(* IEC 61131-3 sources: daoli-st-library/DL_Device (part 12) *)

(* ---- FB_DL_AnalogTransmitter.st ---- *)
(*==============================================================================
 * 组件名称 (Component)  : FB_DL_AnalogTransmitter
 * 所属子库 (Sublibrary) : DL_Device
 * 当前版本 (Version)    : 1.0.0
 * 兼容性   (Platform)   : CODESYS 3.5 / TwinCAT 3 / 汇川 InoProShop / Machine Expert
 *                         仅依赖 Standard.library，零厂商方言
 * 分类     (Category)   : 设备信号处理功能块（Function Block，实现 I_DL_AnalogSensor）
 * 功能简述 (Function)   : NAMUR NE43 语义模拟量变送器处理块。在原始物理域
 *                         （mA/0..10V，由调用方约定）执行四段诊断：故障门限外
 *                         断线（方向可配置）、欠量程段、有效测量域、超量程段，
 *                         0 域附近判回路开路；内嵌滑动平均滤波与线性标定；
 *                         故障态保持末次有效工程量；HH/H/L/LL 四级报警在
 *                         有效与欠/超量程段照常计算、故障态全部保持。
 * 接口实现 (Implements) : I_DL_AnalogSensor（属性 fValue/eQuality/bAlarmHH/
 *                         bAlarmH/bAlarmL/bAlarmLL/uErrorId，全部在本文件
 *                         尾部落地）
 * 开源溯源 (Origin)     : 来源标签 namur-ne43（RAW_NOTES_R5 S-5：NAMUR NE43
 *                         信号电平域，公开推荐实践，多来源交叉印证——有效
 *                         测量域 3.8~20.5 mA、故障域 <3.6 / >21 mA、0 mA =
 *                         回路断线、断线诊断须在原始域而非工程量域判定、
 *                         故障方向可配置、超量程标记而非剔除；仅借鉴公开
 *                         标准语义，欠/超量程段以故障门限与量程端点为界
 *                         （默认 4~20 mA 组态下对应 NE43 3.8/20.5 mA 有效
 *                         域界语义），不硬编码，clean-room 未复制任何源码行）。
 * 红线自检 (Redline)    : R1 零全局变量表/外部变量引用 ✓｜R2 零物理 IO 地址 ✓
 *                         R3 纯 IEC 61131-3 ✓｜R4 防除零/防越界/NaN 自比防御 ✓
 *                         R5 全变量中英双语同行注释 ✓｜R6 质量分级判定含
 *                         ELSE 兜底链 ✓｜R7 滤波实例主体无条件刷新（无定时
 *                         器/边缘实例，滤波为纯算术递推）✓
 * 公约遵循 (Convention) : 0.1 首扫判据 IF bTrack OR (NOT _bInit)，跟踪脉冲
 *                         运行中途插入时重置滤波缓冲与保持值。
 *                         0.6 量程对调自修复：对调后继续计算不中断。
 *                         0.8 全部 REAL 输入 fX <> fX 检测，默认值先赋。
 *                         0.7 故障码段位 16#0003_xxxx：【故障级】0003_0210
 *                         NE43 故障态（断线/开路/非有限输入，R15 锁存语义
 *                         由质量位持续标注，原始恢复后自动解除并保持值
 *                         重新跟随）；【信息级】0003_0102 量程对调自修复 /
 *                         0003_0103 欠/超量程提示 / 0003_0104 原始量程跨度
 *                         退化回退（仅写 uErrorId，不设任何故障位，0.2）。
 * 偏离留档 (Deviation)  : 依 R11 头注释留档，共 4 条：
 *                         ① fFilterTC 已按规格 1.6 定稿删除，由 uFilterWindow
 *                           : USINT := 8 滑动平均窗口替代（规格内定稿）。
 *                         ② 引脚表未列 bTrack，为落实 0.1 首扫/跟踪范式与
 *                           "运行中途插入跟踪脉冲"验收向量新增 IN 引脚。
 *                         ③ FC_DL_LinearScale / FB_DL_MovingAverage 本轮
 *                           尚未入库，标定与滤波在本文件内联等价实现（含
 *                           防除零与窗口钳位），两件入库后可无缝外移。
 *                         ④ 对调自修复码 0.6 原文为 16#0001_0001，依 0.7
 *                           段位分配 DL_Device 族取信息级 0003_0102；新增
 *                           0003_0103/0003_0104 按 0.7 之 01xx 信息段顺延。
 * 修订历史 (Revision)   :
 *   2026-11-15  v1.0.0  首版入库（R5 轮 · DL_Device 开库）
 *============================================================================*)

(*-----------------------------------------------------------------------------
 * 枚举: E_DL_BreakDir（归属 FB_DL_AnalogTransmitter，与其同文件）
 * 含义: 断线故障方向配置，由变送器实际 Downscale/Upscale 组态决定；
 *       只判配置方向，另一方向的越限不误报为断线（S-5 提取点②）。
 *----------------------------------------------------------------------------*)
TYPE E_DL_BreakDir :
(
    eLow  := 0,    // 低断方向（Downscale）：原始值低于故障下门限判断线 / Downscale direction, raw below low fault threshold means wire break
    eHigh := 1     // 高断方向（Upscale）：原始值高于故障上门限判断线 / Upscale direction, raw above high fault threshold means wire break
) USINT;
END_TYPE

(*==============================================================================
 * 功能块主体
 *============================================================================*)
FUNCTION_BLOCK FB_DL_AnalogTransmitter IMPLEMENTS I_DL_AnalogSensor
VAR_INPUT
    fRawInput      : REAL;              // 原始输入（Raw input），已线性化的 mA/0..10V 物理域值，单位由调用方约定 / Raw physical-domain input, unit per caller config
    fRawLow        : REAL;              // 原始域量程下限（Raw span low），如 4.0 mA；对调自修复 / Raw span low endpoint, swap self-repair
    fRawHigh       : REAL;              // 原始域量程上限（Raw span high），如 20.0 mA；对调自修复 / Raw span high endpoint, swap self-repair
    fEuLow         : REAL;              // 工程量程下限（Engineering span low），如 0.0 [%] 或 [kPa] / Engineering span low endpoint
    fEuHigh        : REAL;              // 工程量程上限（Engineering span high），如 100.0 [%] 或 [kPa] / Engineering span high endpoint
    eBreakDirection: E_DL_BreakDir := E_DL_BreakDir.eLow; // 断线故障方向（Break direction），eLow=低断 / eHigh=高通，按变送器组态 / Break direction per transmitter config
    fFaultLow      : REAL := 3.6;       // NE43 故障下门限（NE43 low fault threshold），默认 3.6（原始域）/ Low fault threshold in raw domain
    fFaultHigh     : REAL := 21.0;      // NE43 故障上门限（NE43 high fault threshold），默认 21.0（原始域）/ High fault threshold in raw domain
    uFilterWindow  : USINT := 8;        // 滑动平均窗口（Moving-average window），规格定稿替代时间常数引脚，1=直通 / Moving-average window, 1 = pass-through
    bEnableFilter  : BOOL := TRUE;      // 使能滑动平均滤波（Enable moving-average filter），FALSE=直通 / FALSE bypasses filtering
    fAlarmHH       : REAL;              // 上上限报警门限（High-high alarm limit），量纲=工程量 / High-high limit in engineering unit, 非数=禁用 / NaN disables
    fAlarmH        : REAL;              // 上限报警门限（High alarm limit），量纲=工程量，非数=禁用 / High limit in engineering unit, NaN disables
    fAlarmL        : REAL;              // 下限报警门限（Low alarm limit），量纲=工程量，非数=禁用 / Low limit in engineering unit, NaN disables
    fAlarmLL       : REAL;              // 下下限报警门限（Low-low alarm limit），量纲=工程量，非数=禁用 / Low-low limit in engineering unit, NaN disables
    bTrack         : BOOL;              // 跟踪脉冲（Track pulse），上升语义电平：TRUE 拍重置滤波与保持值（R11 偏离新增，见头注释②）/ Track pulse re-primes filter and hold value
END_VAR

VAR_OUTPUT
    fValue         : REAL;              // 工程量当前值（Current engineering value），故障态保持末次有效值 / Holds last good value in fault
    eQuality       : E_DL_SignalQuality; // 信号质量分级（Signal quality grade），NE43 四段诊断 / NE43 diagnostic grade
    bAlarmHH       : BOOL;              // 上上限报警（High-high alarm），有效及欠/超量程段照常计算 / Computed in good and range-violation segments
    bAlarmH        : BOOL;              // 上限报警（High alarm）/ High alarm
    bAlarmL        : BOOL;              // 下限报警（Low alarm）/ Low alarm
    bAlarmLL       : BOOL;              // 下下限报警（Low-low alarm）/ Low-low alarm
    uErrorId       : UDINT;             // 末次故障码（Last error code），0=无故障，段位 16#0003_xxxx / Last error code, 0 = none
    bWireBreak     : BOOL;              // 断线/开路合并位（Wire break merged flag），含开路 / TRUE on wire break or open loop
    bRangeViol     : BOOL;              // 欠/超量程合并位（Range violation merged flag）/ TRUE on under-range or over-range
END_VAR

VAR
    _bInit         : BOOL := FALSE;     // 首扫初始化标志（First-scan init flag），R19 范式判据成员 / R19 paradigm member
    _fHoldEu       : REAL := 0.0;       // 末次有效工程量（Last good engineering value），保持语义载体 / Hold-semantics carrier
    _fValueOut     : REAL := 0.0;       // 输出镜像寄存（Output mirror register），属性与引脚同源 / Mirror shared by pin and property
    _eQualityInt   : E_DL_SignalQuality := E_DL_SignalQuality.eGood; // 质量分级内部寄存（Internal quality register）/ Internal quality register
    _bAlarmHH      : BOOL;              // 上上限报警内部寄存（Internal high-high alarm register）/ Internal alarm register
    _bAlarmH       : BOOL;              // 上限报警内部寄存（Internal high alarm register）/ Internal alarm register
    _bAlarmL       : BOOL;              // 下限报警内部寄存（Internal low alarm register）/ Internal alarm register
    _bAlarmLL      : BOOL;              // 下下限报警内部寄存（Internal low-low alarm register）/ Internal alarm register
    _uErrorIdInt   : UDINT := 0;        // 故障码内部寄存（Internal error code register）/ Internal error code register
    _bFaultState   : BOOL;              // NE43 故障态标志（NE43 fault state flag），断线/开路/非有限输入 / Fault state on break, open loop or non-finite input
    _fRawLoEff     : REAL;              // 对调修复后量程下限（Repaired span low）/ Repaired raw span low endpoint
    _fRawHiEff     : REAL;              // 对调修复后量程上限（Repaired span high）/ Repaired raw span high endpoint
    _bSwap         : BOOL;              // 本拍发生对调修复（Swap repair occurred this cycle）/ Swap repair occurred flag
    _bSpanDegenerate : BOOL;            // 原始量程跨度退化（Degenerate raw span），近零或非有限 / Span near zero or non-finite
    _fFaultLoEff   : REAL := 3.6;       // 防御后故障下门限（Sanitized low fault threshold）/ Sanitized low fault threshold
    _fFaultHiEff   : REAL := 21.0;      // 防御后故障上门限（Sanitized high fault threshold）/ Sanitized high fault threshold
    _fEuLoEff      : REAL := 0.0;       // 防御后工程下限（Sanitized engineering low）/ Sanitized engineering low
    _fEuHiEff      : REAL := 100.0;     // 防御后工程上限（Sanitized engineering high）/ Sanitized engineering high
    _bValid        : BOOL;              // 原始输入有效（Raw input valid），非有限值为 FALSE / FALSE when input is non-finite
    _fScaleRaw     : REAL;              // 参与标定的原始值（Raw value entering scaling），滤波输出或直通 / Filtered or pass-through raw value
    _fScaledEu     : REAL;              // 本拍标定结果（Scaled result this cycle）/ Scaled engineering result this cycle
    _fRawSpan      : REAL;              // 原始量程跨度（Raw span width）/ Raw span width
    _bFilterActive : BOOL;              // 滤波激活（Filter active），使能且窗口 >= 2 / Active when enabled and window >= 2
    _uWindowEff    : USINT;             // 钳位后有效窗口（Effective clamped window），上限 128 / Effective window clamped to 128
    _uWindowPrev   : USINT;             // 上一拍有效窗口（Previous effective window），变更检测用于缓冲重置 / Previous window for change detection
    _uBufIdx       : UINT;              // 环形缓冲写指针（Ring buffer write index），0..127 / Ring write index 0..127
    _uBufFill      : USINT;             // 有效样本数（Valid sample count），上限=有效窗口 / Valid samples, capped at effective window
    _fBufSum       : REAL := 0.0;       // 窗口样本和（Window sample sum），每拍重算 / Recomputed each cycle
    _fFillR        : REAL := 1.0;       // 样本数实型镜像（Sample count REAL mirror），供安全除法 / REAL mirror of sample count for safe division
    _afBuf         : ARRAY[0..127] OF REAL; // 滑动平均环形缓冲（Moving-average ring buffer），128 槽 / 128-slot ring buffer
    i              : UINT;              // 缓冲遍历循环索引（Buffer traversal loop index）/ Loop index for buffer traversal
    _uRingIdx      : UINT;              // 环形取数临时索引（Ring fetch temp index）/ Temporary ring fetch index
END_VAR

// ============================================================================
// 段 1｜首扫/跟踪初始化（R19 唯一合法范式：IF bTrack OR (NOT _bInit)）
//      First-scan / track initialization (R19 sole legal paradigm)
// ============================================================================
IF bTrack OR (NOT _bInit) THEN
    _uBufIdx   := 0;                          // 写指针归零（Write index reset）
    _uBufFill  := 0;                          // 有效样本清零：滤液从直通逐步重新填充（Samples cleared, filter refills from pass-through）
    _fBufSum   := 0.0;                        // 窗口和清零（Window sum cleared）
    _fHoldEu   := 0.0;                        // 保持值清零，本拍有效样本将立即回填（Hold cleared, refilled by first valid sample）
    _bFaultState := FALSE;                    // 故障态复位（Fault state released）
    _uErrorIdInt := 0;                        // 故障码清零（Error code cleared）
    _eQualityInt := E_DL_SignalQuality.eGood; // 质量复位为良好（Quality reset to good）
    _bInit      := TRUE;                      // 初始化完成（Initialization done）
END_IF

// ============================================================================
// 段 2｜窗口参数钳位与变更检测（防越界：窗口上限 128 槽缓冲）
//      Window clamping and change detection (bounds defense: 128-slot buffer)
// ============================================================================
_uWindowEff := uFilterWindow;                 // 取组态窗口（Take configured window）
IF _uWindowEff > 128 THEN
    _uWindowEff := 128;                       // 超限钳位到缓冲容量（Clamp to buffer capacity）
END_IF
IF _uWindowEff = 0 THEN
    _uWindowEff := 1;                         // 零窗口按单样本直通（Zero window treated as single-sample pass-through）
END_IF
IF _uWindowEff <> _uWindowPrev THEN           // 窗口在线变更（Window changed online）
    _uBufFill := 0;                           // 缓冲判无效重新填充（Invalidate buffer, refill from scratch）
    _uWindowPrev := _uWindowEff;              // 记录新窗口（Record new window）
END_IF
_bFilterActive := bEnableFilter AND (_uWindowEff >= 2); // 窗口 1 视为直通（Window 1 treated as pass-through）

// ============================================================================
// 段 3｜参数防御（0.8：全部 REAL 参数先做非数自比，默认值先赋）+ 0.6 对调自修复
//      Parameter sanitation (0.8 NaN self-compare, defaults first) + 0.6 swap repair
// ============================================================================
_fRawLoEff := fRawLow;                        // 量程下限镜像（Span low mirror）
_fRawHiEff := fRawHigh;                       // 量程上限镜像（Span high mirror）
_fEuLoEff  := fEuLow;                         // 工程下限镜像（Engineering low mirror）
_fEuHiEff  := fEuHigh;                        // 工程上限镜像（Engineering high mirror）
_fFaultLoEff := fFaultLow;                    // 故障下门限镜像（Low fault threshold mirror）
_fFaultHiEff := fFaultHigh;                   // 故障上门限镜像（High fault threshold mirror）

IF _fFaultLoEff <> _fFaultLoEff THEN          // 非数自比检测（NaN self-compare test）
    _fFaultLoEff := 3.6;                      // 回落 NE43 默认下门限（Fallback to NE43 default low）
END_IF
IF _fFaultHiEff <> _fFaultHiEff THEN          // 非数自比检测（NaN self-compare test）
    _fFaultHiEff := 21.0;                     // 回落 NE43 默认上门限（Fallback to NE43 default high）
END_IF
IF _fEuLoEff <> _fEuLoEff THEN                // 非数自比检测（NaN self-compare test）
    _fEuLoEff := 0.0;                         // 回落工程下限默认（Fallback engineering low default）
END_IF
IF _fEuHiEff <> _fEuHiEff THEN                // 非数自比检测（NaN self-compare test）
    _fEuHiEff := 100.0;                       // 回落工程上限默认（Fallback engineering high default）
END_IF

_bSwap := FALSE;                              // 对调标志复位（Swap flag reset）
IF _fRawLoEff > _fRawHiEff THEN               // 参数对自修复判据（Pair swap test, NaN-safe ordering）
    _fRawLoEff := fRawHigh;                   // 下限取原上限（Low takes former high）
    _fRawHiEff := fRawLow;                    // 上限取原下限（High takes former low）
    _bSwap := TRUE;                           // 登记对调修复（Register swap repair, computation continues）
END_IF

// ============================================================================
// 段 4｜非有限输入判定（0.8）与出口默认值先赋（保持语义）
//      Non-finite input test (0.8) and output defaults assigned first (hold)
// ============================================================================
_bValid := (fRawInput = fRawInput);           // 非数自比检测：等号成立即有效（NaN 时自比不等）/ NaN iff self-compare fails, TRUE means valid
_fValueOut := _fHoldEu;                       // 出口默认：保持末次有效值（Default: hold last good value）
_bFaultState := FALSE;                        // 故障态先复位，分级链中重新判定（Fault state preset FALSE, re-decided below）
_eQualityInt := E_DL_SignalQuality.eGood;     // 出口默认质量（Default quality）

// ============================================================================
// 段 5｜NE43 四段质量分级（全部在原始物理域判定，S-5 提取点③；
//       断线只判配置方向，配置外方向不误报）
//      NE43 four-band classification in raw domain, break judged only on
//      the configured direction to avoid false breaks
// ============================================================================

IF NOT _bValid THEN
    _eQualityInt := E_DL_SignalQuality.eOpenLoop;   // 非有限输入按回路开路处理（Non-finite input as open loop）
    _bFaultState := TRUE;                           // 进入故障态（Enter fault state）
ELSIF fRawInput < (_fFaultLoEff * 0.5) THEN
    _eQualityInt := E_DL_SignalQuality.eOpenLoop;   // 0 域附近判开路（0 mA 回路断开）/ Near-zero domain as open loop
    _bFaultState := TRUE;
ELSIF fRawInput < _fFaultLoEff THEN
    IF eBreakDirection = E_DL_BreakDir.eLow THEN
        _eQualityInt := E_DL_SignalQuality.eWireBreakLow; // 配置低断：判断线（Configured downscale: wire break）
        _bFaultState := TRUE;
    ELSE
        _eQualityInt := E_DL_SignalQuality.eUnderRange;   // 配置高通：欠量程段不误报断线（High config: under-range, no false break）
    END_IF
ELSIF fRawInput > _fFaultHiEff THEN
    IF eBreakDirection = E_DL_BreakDir.eHigh THEN
        _eQualityInt := E_DL_SignalQuality.eWireBreakHigh; // 配置高通：判断线（Configured upscale: wire break）
        _bFaultState := TRUE;
    ELSE
        _eQualityInt := E_DL_SignalQuality.eOverRange;     // 配置低断：超量程段不误报断线（Low config: over-range, no false break）
    END_IF
ELSIF fRawInput < _fRawLoEff THEN
    _eQualityInt := E_DL_SignalQuality.eUnderRange;   // 欠量程段（如 3.6~4.0 mA）标记不剔除（Under-range marked, not discarded）
ELSIF fRawInput > _fRawHiEff THEN
    _eQualityInt := E_DL_SignalQuality.eOverRange;    // 超量程段（如 20.0~21.0 mA）标记不剔除（Over-range marked, not discarded）
ELSE
    _eQualityInt := E_DL_SignalQuality.eGood;         // 有效测量域（Valid measurement span）
END_IF

// ============================================================================
// 段 6｜滑动平均滤波（仅有效拍推入缓冲，故障拍不污染窗口）+ 线性标定
//      Moving-average filter (push only on valid cycles) + linear scaling
// ============================================================================
IF _bFaultState THEN
    _fScaleRaw := fRawInput;                  // 故障拍标定值不使用（Unused in fault cycles, hold applies）
ELSE
    IF _bFilterActive THEN
        _afBuf[_uBufIdx] := fRawInput;        // 写入环形槽（Write ring slot, index < 128 by MOD）
        _uBufIdx := (_uBufIdx + 1) MOD 128;   // 写指针循环推进（Advance write index cyclically）
        IF _uBufFill < _uWindowEff THEN
            _uBufFill := _uBufFill + 1;       // 未满则递增有效样本（Increment fill until window reached）
        END_IF
        _fBufSum := 0.0;                      // 每拍重算窗口和（Recompute window sum each cycle）
        FOR i := 1 TO _uBufFill DO            // 固定界循环，无死循环风险（Bounded loop, no deadlock risk）
            _uRingIdx := (_uBufIdx + 128 - i) MOD 128; // 倒序取最近样本槽（Fetch latest slots in reverse order）
            _fBufSum := _fBufSum + _afBuf[_uRingIdx];  // 累加窗口样本（Accumulate window sample）
        END_FOR
        _fFillR := _uBufFill;                 // 样本数实型镜像（Sample count as REAL）
        IF _fFillR > 0.5 THEN
            _fScaleRaw := _fBufSum / _fFillR; // 窗口均值（Window mean, divisor proven >= 1）
        ELSE
            _fScaleRaw := fRawInput;          // 防除零回退直通（Divide-by-zero fallback to pass-through）
        END_IF
    ELSE
        _fScaleRaw := fRawInput;              // 滤波禁用直通（Filter disabled, pass-through）
    END_IF

    // 线性标定（内联实现，偏离留档③；除零与退化双重防御）
    _fRawSpan := _fRawHiEff - _fRawLoEff;     // 原始量程跨度（Raw span width）
    _bSpanDegenerate := (_fRawSpan <> _fRawSpan) OR (ABS(_fRawSpan) < 1E-9); // 非数或近零判退化（Degenerate on NaN or near-zero）
    IF _bSpanDegenerate THEN
        _fScaledEu := _fEuLoEff;              // 退化回退工程下限（Degenerate fallback to engineering low）
    ELSE
        _fScaledEu := _fEuLoEff + (_fScaleRaw - _fRawLoEff) * (_fEuHiEff - _fEuLoEff) / _fRawSpan; // 线性插值（Linear interpolation, denominator proven non-zero）
    END_IF
    _fValueOut := _fScaledEu;                 // 有效拍输出跟随（Output follows on valid cycles）
    _fHoldEu   := _fScaledEu;                 // 更新保持载体（Update hold carrier）
END_IF

// ============================================================================
// 段 7｜四级报警计算（有效与欠/超量程段照常计算；故障态全部保持；
//       门限为非数时该级视为未组态不报警——0.8 防御）
//      Four-level alarms (computed in good and range segments, held in
//      fault; NaN threshold disables that level)
// ============================================================================
IF NOT _bFaultState THEN
    IF fAlarmHH = fAlarmHH THEN
        _bAlarmHH := (_fValueOut >= fAlarmHH); // 上上限判定（High-high evaluation）
    ELSE
        _bAlarmHH := FALSE;                    // 门限非数=该级禁用（NaN limit disables level）
    END_IF
    IF fAlarmH = fAlarmH THEN
        _bAlarmH := (_fValueOut >= fAlarmH);   // 上限判定（High evaluation）
    ELSE
        _bAlarmH := FALSE;                     // 门限非数=该级禁用（NaN limit disables level）
    END_IF
    IF fAlarmL = fAlarmL THEN
        _bAlarmL := (_fValueOut <= fAlarmL);   // 下限判定（Low evaluation）
    ELSE
        _bAlarmL := FALSE;                     // 门限非数=该级禁用（NaN limit disables level）
    END_IF
    IF fAlarmLL = fAlarmLL THEN
        _bAlarmLL := (_fValueOut <= fAlarmLL); // 下下限判定（Low-low evaluation）
    ELSE
        _bAlarmLL := FALSE;                    // 门限非数=该级禁用（NaN limit disables level）
    END_IF
END_IF // 故障态不进入本段，四级报警输出自动保持上一拍值（Fault cycles skip this block, alarms held）

// ============================================================================
// 段 8｜故障码优先级链与合并位派生（信息级仅写 uErrorId，0.2 公约）
//      Error-code priority chain and merged flag derivation (info codes only)
// ============================================================================
IF _bFaultState THEN
    _uErrorIdInt := 16#0003_0210;             // 0003_0210 NE43 故障态（断线/开路/非有限输入）【故障级】/ NE43 fault state, fault level
ELSIF (_eQualityInt = E_DL_SignalQuality.eUnderRange) OR (_eQualityInt = E_DL_SignalQuality.eOverRange) THEN
    _uErrorIdInt := 16#0003_0103;             // 0003_0103 欠/超量程提示【信息级】/ Range violation hint, info level
ELSIF _bSwap THEN
    _uErrorIdInt := 16#0003_0102;             // 0003_0102 量程对调自修复【信息级】（0.6 公约，段位依 0.7 归 DL_Device 信息段）/ Swap self-repair, info level
ELSIF _bSpanDegenerate THEN
    _uErrorIdInt := 16#0003_0104;             // 0003_0104 原始量程跨度退化回退【信息级】/ Degenerate span fallback, info level
ELSE
    _uErrorIdInt := 0;                        // 无故障无提示（No fault, no hint）
END_IF

// ============================================================================
// 段 9｜引脚映射（属性与引脚同源于内部镜像，避免同名遮蔽）
//      Pin mapping (pin and property share internal mirrors, no shadowing)
// ============================================================================
fValue     := _fValueOut;                     // 工程量输出（Engineering value output）
eQuality   := _eQualityInt;                   // 质量分级输出（Quality output）
bAlarmHH   := _bAlarmHH;                      // 上上限输出（High-high output）
bAlarmH    := _bAlarmH;                       // 上限输出（High output）
bAlarmL    := _bAlarmL;                       // 下限输出（Low output）
bAlarmLL   := _bAlarmLL;                      // 下下限输出（Low-low output）
uErrorId   := _uErrorIdInt;                   // 故障码输出（Error code output）
bWireBreak := (_eQualityInt = E_DL_SignalQuality.eWireBreakLow)
          OR (_eQualityInt = E_DL_SignalQuality.eWireBreakHigh)
          OR (_eQualityInt = E_DL_SignalQuality.eOpenLoop);            // 断线/开路合并位（Break/open merged flag）
bRangeViol := (_eQualityInt = E_DL_SignalQuality.eUnderRange)
          OR (_eQualityInt = E_DL_SignalQuality.eOverRange);           // 欠/超量程合并位（Range violation merged flag）

(*------------------------------------------------------------------------------
 * 属性: fValue（GET）—— 工程量当前值（故障态保持末次有效值）。
 *      Property fValue (GET) - current engineering value, holds last good in fault.
 *------------------------------------------------------------------------------*)
PROPERTY fValue : REAL
fValue := _fValueOut;         // 返回输出镜像（Return output mirror）

(*------------------------------------------------------------------------------
 * 属性: eQuality（GET）—— 信号质量分级（NE43 四段诊断结果）。
 *      Property eQuality (GET) - signal quality grade per NE43 diagnostics.
 *------------------------------------------------------------------------------*)
PROPERTY eQuality : E_DL_SignalQuality
eQuality := _eQualityInt;     // 返回质量镜像（Return quality mirror）

(*------------------------------------------------------------------------------
 * 属性: bAlarmHH（GET）—— 上上限报警位。
 *      Property bAlarmHH (GET) - high-high alarm bit.
 *------------------------------------------------------------------------------*)
PROPERTY bAlarmHH : BOOL
bAlarmHH := _bAlarmHH;        // 返回上上限镜像（Return high-high mirror）

(*------------------------------------------------------------------------------
 * 属性: bAlarmH（GET）—— 上限报警位。
 *      Property bAlarmH (GET) - high alarm bit.
 *------------------------------------------------------------------------------*)
PROPERTY bAlarmH : BOOL
bAlarmH := _bAlarmH;          // 返回上限镜像（Return high mirror）

(*------------------------------------------------------------------------------
 * 属性: bAlarmL（GET）—— 下限报警位。
 *      Property bAlarmL (GET) - low alarm bit.
 *------------------------------------------------------------------------------*)
PROPERTY bAlarmL : BOOL
bAlarmL := _bAlarmL;          // 返回下限镜像（Return low mirror）

(*------------------------------------------------------------------------------
 * 属性: bAlarmLL（GET）—— 下下限报警位。
 *      Property bAlarmLL (GET) - low-low alarm bit.
 *------------------------------------------------------------------------------*)
PROPERTY bAlarmLL : BOOL
bAlarmLL := _bAlarmLL;        // 返回下下限镜像（Return low-low mirror）

(*------------------------------------------------------------------------------
 * 属性: uErrorId（GET）—— 末次故障码（0=无故障）。
 *      Property uErrorId (GET) - last error code (0 = none).
 *------------------------------------------------------------------------------*)
PROPERTY uErrorId : UDINT
uErrorId := _uErrorIdInt;     // 返回故障码镜像（Return error code mirror）
END_FUNCTION_BLOCK

(* ---- FB_DL_AnalogValve.st ---- *)
(*==============================================================================
 * 组件名称 (Component)  : FB_DL_AnalogValve
 * 所属子库 (Sublibrary) : DL_Device
 * 当前版本 (Version)    : 1.0.1
 * 兼容性   (Platform)   : CODESYS 3.5 / TwinCAT 3 / 汇川 InoProShop / Machine Expert
 *                         仅依赖 Standard.library（TON / R_TRIG），零厂商方言
 * 分类     (Category)   : 设备执行器功能块（Function Block，实现 I_DL_ProportionalValve）
 * 功能简述 (Function)   : 模拟量比例阀指令整形与诊断功能块（不含阀位闭环，
 *                         闭环由驱动器/上层 PID 完成，本块职责单一）。
 *                         透传+补偿链：设定钳位 [0,100] → 零点死区补偿
 *                         （防阀芯微抖）→ 限幅域映射 → 阀位指令输出；
 *                         偏差报警延时确认（瞬时型每拍重算，恢复自动清）；
 *                         非有限值反馈锁存保持末次有效值；限幅域对调
 *                         自修复；状态机 E_DL_ValveState + CASE + ELSE
 *                         兜底。
 * 接口实现 (Implements) : I_DL_ProportionalValve。接口 OUT 列同名成员
 *                         （eState/fPosCmd/fPosFeedback/bDeviationAlarm/
 *                         bFault/uErrorId）按 R22 以只读 PROPERTY GET
 *                         承载（内部镜像同源；fPosFeedback 为 IN 引脚与
 *                         接口属性双形式暴露，沿用库级既有先例），非接口
 *                         成员 fPosOutput 保留 VAR_OUTPUT；方法
 *                         SetPosition/CmdStop/CmdReset 全部在本文件尾部
 *                         落地。
 * 开源溯源 (Origin)     : 来源标签 lbp-basic-process / lbp-device
 *                         （RAW_NOTES_R6 S-1：比例阀指令整形链（钳位-死区
 *                         补偿-限幅域映射）、偏差延时报警、限幅域端点组态
 *                         等行业公知工程惯例，公开教学资料，仅借鉴通用
 *                         工程语义；状态机、整形链实现、故障码按本库红线
 *                         独立设计，clean-room 未复制源码）。
 * 红线自检 (Redline)    : R1 零全局变量表/外部变量引用 ✓｜R2 零物理 IO 地址 ✓
 *                         R3 纯 IEC 61131-3 ✓｜R4 防除零/防越界/非有限值
 *                         防御/浮点容差比较 ✓｜R5 全变量中英双语同行注释 ✓
 *                         R6 ENUM+CASE+ELSE ✓｜R7 两个定时器/边缘实例主体
 *                         最前部无条件刷新 ✓
 * 公约遵循 (Convention) : 0.1/R23 本块为逐拍组合整形链（设定→钳位→死区→
 *                         映射，全部由实时输入重算自校正），无积分/滤波类
 *                         需要首扫初始化的连续量驻留状态，免首扫（无
 *                         bInit 标志）；时间基准按公约 0.5 采用 TON 延时
 *                         引脚（偏差确认），无采样周期类连续量语义。
 *                         0.6 限幅域对调自修复：fOutMin > fOutMax 时对调
 *                         + 置信息级码 + 继续计算不中断。
 *                         0.7 故障码段位 16#0003_xxxx：【故障级】0003_0260
 *                         阀位反馈信号无效 / 0003_0261 非法状态，R15 锁存
 *                         仅复位可清；【信息级】0003_0108 设定值钳位 /
 *                         0003_0109 输出限幅域对调自修复 / 0003_0112 偏差
 *                         报警激活（瞬时型每拍重算，0.15；不进 bFault）。
 * 偏离留档 (Deviation)  : 依 R11 头注释留档，共 1 条：
 *                         ① 信息级码：规格原分配 0003_0105/0106，经与子库
 *                           VERSION.md 故障码表核对，R5 已占用 0102~0104
 *                           （AnalogTransmitter），且 0106/0107 已由本轮
 *                           变频器块顺延占用（0105 经终审裁定空置：重启抑
 *                           制拒绝统一沿用 DolMotor 既有语义码位 0208），
 *                           依公约 0.7 冲突顺延：设定值钳位 → 0108、限幅
 *                           域对调 → 0109；偏差报警激活为新码位，顺延分配
 *                           0112。
 * 修订历史 (Revision)   :
 *   2026-11-15  v1.0.0  首版入库（R6 轮 · DL_Device 阀门/驱动族深化）
 *   2026-11-15  v1.0.1  终审修复【工程语义级】限幅域对调穿透：原实现对调时
 *                       直读原始引脚（fOutMin/fOutMax），混合非数组态下
 *                       （如下端非数+上端负值）会把未防御的 NaN 带回生效
 *                       域并经映射链输出 NaN 阀位指令且不带故障码。修法：
 *                       对调改为经中间变量交换已防御的生效值。引脚契约
 *                       零变更。
 *============================================================================*)
FUNCTION_BLOCK FB_DL_AnalogValve IMPLEMENTS I_DL_ProportionalValve
VAR_INPUT
    fPosSetpoint     : REAL;            // 阀位设定（Position setpoint）[%]，0..100，越界钳位信息级 / Position setpoint [%], clamped with info code
    fPosFeedback     : REAL;            // 阀位反馈（Position feedback）[%]，0..100，来自阀位变送器；非有限值防御 / Position feedback [%] from transmitter, non-finite defended
    fZeroDeadband    : REAL := 0.5;     // 零点死区补偿（Zero deadband compensation）[%]，输出小于此值钳为 0 防阀芯微抖 / Zero deadband [%], output below clamped to zero
    fDeviationLimit  : REAL := 5.0;     // 偏差报警门限（Deviation limit）[%]，默认 5.0 / Deviation alarm limit [%], default 5.0
    tDeviationDelay  : TIME := T#10S;   // 偏差报警确认延时（Deviation delay），防动态调节过程误报 / Deviation confirmation delay against dynamic transients
    fOutMin          : REAL := 0.0;     // 输出限幅域下端点（Output span low endpoint）[%]，对调自修复 / Output span low endpoint, swap self-repair
    fOutMax          : REAL := 100.0;   // 输出限幅域上端点（Output span high endpoint）[%]，对调自修复 / Output span high endpoint, swap self-repair
    bEnable          : BOOL;            // 调节使能（Modulating enable），FALSE 时输出冻结保持 / Modulating enable, FALSE freezes output hold
    bReset           : BOOL;            // 故障复位（Fault reset），上升沿生效 / Fault reset, rising edge effective
END_VAR

VAR_OUTPUT
    fPosOutput : REAL;                  // 阀位指令输出（Position output）[%]，死区补偿+限幅域映射后，量纲=限幅域（R20）/ Shaped position output [%], span of limit domain
END_VAR

VAR
    _eState        : E_DL_ValveState := E_DL_ValveState.eIdle; // 内部状态机步序（Internal state step），外部经属性只读 / Internal state, read-only via property
    _bFaultLatch   : BOOL;              // 故障锁存标志（Fault latch flag），仅复位清除 / Fault latch flag, cleared only by reset
    _uErrorIdInt   : UDINT;             // 故障级码内部寄存（Internal fault-code register） / Internal fault-level code register
    _uInfoCode     : UDINT;             // 本拍信息级码（Info code this cycle），瞬时型每拍重算（0.15）/ Transient info code recomputed each cycle
    _bHoldLatch    : BOOL;              // 输出冻结锁存（Output freeze latch），CmdStop 置位 / Output freeze latch set by CmdStop
    _bPendReset    : BOOL;              // 方法复位请求（Method reset request），由 CmdReset 置位 / Method reset request set by CmdReset
    _bClampOccur   : BOOL;              // 本拍设定值钳位发生（Setpoint clamp occurred this cycle）/ Setpoint clamp occurred flag
    _fPosMethVal   : REAL;              // 方法阀位设定值（Method position value）[%] / Position value set via method
    _bPosMethAct   : BOOL;              // 方法阀位设定激活（Method position active），激活后覆盖引脚 / Method position active, overrides pin
    _fPosFbHold    : REAL := 0.0;       // 末次有效阀位反馈（Last valid position feedback）[%]，保持载体 / Last valid feedback hold carrier
    _fPosCmdEff    : REAL := 0.0;       // 钳位+死区后生效阀位指令（Effective command after clamp and deadband）[%] / Effective command [%]
    _fPosOutHold   : REAL := 0.0;       // 输出保持载体（Output hold carrier）[%]，冻结/故障态保持 / Output hold carrier [%]
    _fOutMinEff    : REAL := 0.0;       // 对调修复后限幅域下端（Repaired span low endpoint）[%] / Repaired span low endpoint
    _fOutMaxEff    : REAL := 100.0;     // 对调修复后限幅域上端（Repaired span high endpoint）[%] / Repaired span high endpoint
    _fZeroDbEff    : REAL := 0.5;       // 防御后死区（Sanitized deadband）[%]，非数/负值钳零 / Sanitized deadband, NaN or negative clamped to zero
    _fDevLimEff    : REAL := 5.0;       // 防御后偏差门限（Sanitized deviation limit）[%] / Sanitized deviation limit
    _bSpanSwap     : BOOL;              // 本拍限幅域对调修复（Span swap repair this cycle）/ Span swap repair occurred flag
    _fSpanTmp      : REAL;              // 对调交换中间变量（Swap temp carrier）[%]，生效域已防御值 / Swap temp for sanitized span values
    _bSpanDegenerate : BOOL;            // 限幅域跨度退化（Degenerate span），近零或非有限 / Span degenerate on near-zero or NaN
    _bFbValid      : BOOL;              // 本拍反馈有效性（Feedback validity this cycle），非有限值为 FALSE / FALSE when feedback non-finite
    _bDevRaw       : BOOL;              // 偏差越限原始判据（Raw deviation-exceed test）/ Raw deviation exceed flag
    _bDeviationAct : BOOL;              // 偏差报警激活中（Deviation alarm active），延时确认后 / Deviation alarm active after confirmation delay
    _fbTrigReset   : R_TRIG;            // 引脚复位上升沿（Pin reset edge）/ Pin reset rising edge
    _fbTonDev      : TON;               // 偏差报警确认延时定时器（Deviation confirmation timer）/ Deviation confirmation timer
END_VAR

METHOD SetPosition : BOOL
VAR_INPUT
    fPos : REAL; // 阀位设定值（Position value）[%]，域 0..100 / Position value [%], range 0..100
END_VAR
IF _bFaultLatch OR (_eState = E_DL_ValveState.eFault) THEN
    SetPosition := FALSE;     // 故障态拒绝（Rejected in fault state）
ELSIF (fPos <> fPos) OR (fPos < 0.0) OR (fPos > 100.0) THEN
    SetPosition := FALSE;     // 非数或越域拒绝（Rejected on NaN or out of range）
ELSE
    _fPosMethVal := fPos;     // 登记方法设定值（Register method position value）
    _bPosMethAct := TRUE;     // 激活方法设定通道（Activate method source channel）
    _bHoldLatch  := FALSE;    // 设定即解除输出冻结（Set releases output freeze）
    SetPosition := TRUE;      // 受理成功（Accepted）
END_IF

(*------------------------------------------------------------------------------
 * 方法: CmdStop —— 冻结输出保持当前阀位，直至下次设定或使能撤除。
 *      Method CmdStop - freeze output until next set or enable drop.
 *------------------------------------------------------------------------------*)
    END_METHOD

METHOD CmdStop : BOOL
VAR_INPUT
END_VAR
IF _bFaultLatch OR (_eState = E_DL_ValveState.eFault) THEN
    CmdStop := FALSE;         // 故障态拒绝（Rejected in fault state）
ELSE
    _bHoldLatch := TRUE;      // 登记冻结锁存，主体状态机消化（Register freeze latch, consumed by body）
    CmdStop := TRUE;          // 受理成功（Accepted）
END_IF

(*------------------------------------------------------------------------------
 * 方法: CmdReset —— 复位故障，返回是否可复位（存在锁存故障时为 TRUE）。
 *      Method CmdReset - reset fault, returns TRUE only when a latch exists.
 *------------------------------------------------------------------------------*)
    END_METHOD

METHOD CmdReset : BOOL
VAR_INPUT
END_VAR
IF _bFaultLatch OR (_eState = E_DL_ValveState.eFault) THEN
    _bPendReset := TRUE;      // 登记复位请求，主体状态机消化（Register reset request, consumed by body）
    CmdReset := TRUE;         // 可复位（Resettable）
ELSE
    CmdReset := FALSE;        // 无故障可复位（Nothing to reset）
END_IF

(*------------------------------------------------------------------------------
 * 属性: eState（GET）—— 当前状态机状态只读视图。
 *      Property eState (GET) - read-only view of the current state machine state.
 *------------------------------------------------------------------------------*)
    END_METHOD

// ============================================================================
// 段 1｜定时器与边缘检测实例无条件周期刷新（R7：严禁置于 IF/CASE 分支内）
//      Unconditional per-cycle refresh of all timer and edge instances (R7)
// ============================================================================
_fbTrigReset(CLK := bReset);
_bDevRaw := (_eState = E_DL_ValveState.eModulating) AND (ABS(_fPosCmdEff - _fPosFbHold) > _fDevLimEff); // 偏差原始判据（Raw deviation test）
_fbTonDev(IN := _bDevRaw, PT := tDeviationDelay); // 延时确认防动态调节误报（Delay confirmation against dynamics）

// ============================================================================
// 段 2｜参数防御（0.8：非数自比检测，默认值先赋）+ 0.6 限幅域对调自修复
//      Parameter sanitation (0.8 NaN self-compare) + 0.6 span swap repair
// ============================================================================
_uInfoCode := 0;                      // 本拍信息级码先归零，事件段重算（Info code preset zero, recomputed in event chain）
_bClampOccur := FALSE;                // 钳位标志复位（Clamp flag reset）
_fZeroDbEff := fZeroDeadband;         // 死区镜像（Deadband mirror）
IF _fZeroDbEff <> _fZeroDbEff THEN    // 非数自比检测（NaN self-compare test）
    _fZeroDbEff := 0.0;               // 非数死区钳零禁用补偿（NaN deadband clamped to zero, compensation disabled）
END_IF
IF _fZeroDbEff < 0.0 THEN
    _fZeroDbEff := 0.0;               // 负死区钳零（Negative deadband clamped to zero）
END_IF
_fDevLimEff := fDeviationLimit;       // 偏差门限镜像（Deviation limit mirror）
IF _fDevLimEff <> _fDevLimEff THEN    // 非数自比检测（NaN self-compare test）
    _fDevLimEff := 5.0;               // 回落默认门限（Fallback to default limit）
END_IF
IF _fDevLimEff < 0.0 THEN
    _fDevLimEff := ABS(_fDevLimEff);  // 负门限取绝对值保持报警有效（Negative limit made absolute, alarm stays valid）
END_IF

_fOutMinEff := fOutMin;               // 限幅域下端镜像（Span low mirror）
_fOutMaxEff := fOutMax;               // 限幅域上端镜像（Span high mirror）
IF _fOutMinEff <> _fOutMinEff THEN    // 非数自比检测（NaN self-compare test）
    _fOutMinEff := 0.0;               // 回落下端默认（Fallback to default low）
END_IF
IF _fOutMaxEff <> _fOutMaxEff THEN    // 非数自比检测（NaN self-compare test）
    _fOutMaxEff := 100.0;             // 回落上端默认（Fallback to default high）
END_IF
_bSpanSwap := FALSE;                  // 对调标志复位（Swap flag reset）
IF _fOutMinEff > _fOutMaxEff THEN     // 参数对自修复判据（Pair swap test）
    _fSpanTmp     := _fOutMinEff;     // 对调经已防御的生效值交换（中间变量，防原始引脚
    _fOutMinEff   := _fOutMaxEff;     // 非有限值穿透——若直读原始引脚，混合非数组态
    _fOutMaxEff   := _fSpanTmp;       // 会把 NaN 带回生效域，终审修复）
    _bSpanSwap := TRUE;               // 登记对调修复，继续计算不中断（Register swap repair, computation continues）
END_IF

// ============================================================================
// 段 3｜阀位反馈有效性全局监视（优先级最高，故障级锁存保持末次有效值）
//      Position feedback validity global monitor (highest priority, latched)
// ============================================================================
_bFbValid := (fPosFeedback = fPosFeedback); // 非数自比检测：等号成立即有效（NaN iff self-compare fails）
IF _bFbValid THEN
    _fPosFbHold := fPosFeedback;      // 更新末次有效反馈（Update last valid feedback）
ELSE
    _bFaultLatch := TRUE;             // 反馈失效锁存（Feedback loss latch）
    _uErrorIdInt := 16#0003_0260;     // 0003_0260 阀位反馈信号无效【故障级】/ Position feedback invalid, fault level
    _eState      := E_DL_ValveState.eFault; // 强制故障态（Force fault state）
END_IF

// ============================================================================
// 段 4｜指令整形链：来源选择 → 钳位 [0,100] → 零点死区补偿
//      Command shaping chain: source select → clamp [0,100] → zero deadband
// ============================================================================
IF _bPosMethAct THEN
    _fPosCmdEff := _fPosMethVal;      // 方法设定覆盖引脚（Method value overrides pin）
ELSE
    _fPosCmdEff := fPosSetpoint;      // 引脚设定（Pin setpoint）
END_IF
IF _fPosCmdEff <> _fPosCmdEff THEN    // 非数自比检测（NaN self-compare test）
    _fPosCmdEff := 0.0;               // 非数设定回零（NaN setpoint falls back to zero）
END_IF
IF _fPosCmdEff < 0.0 THEN
    _fPosCmdEff := 0.0;               // 下限钳位（Clamped to low bound）
    _bClampOccur := TRUE;             // 登记钳位事件（Register clamp event）
END_IF
IF _fPosCmdEff > 100.0 THEN
    _fPosCmdEff := 100.0;             // 上限钳位（Clamped to high bound）
    _bClampOccur := TRUE;             // 登记钳位事件（Register clamp event）
END_IF
IF ABS(_fPosCmdEff) < _fZeroDbEff THEN
    _fPosCmdEff := 0.0;               // 零点死区补偿：近零指令钳为 0 防阀芯微抖（Zero deadband: near-zero command clamped to zero）
END_IF

// ============================================================================
// 段 5｜核心状态机（ENUM + CASE，含 ELSE 非法状态兜底）
//      Core state machine (ENUM + CASE with ELSE illegal-state fallback)
// ============================================================================
IF _bFaultLatch OR (_eState = E_DL_ValveState.eFault) THEN
    CASE _eState OF
        E_DL_ValveState.eFault: // 故障锁存态：输出冻结保持，仅复位可退出
            IF _fbTrigReset.Q OR _bPendReset THEN
                _bPendReset  := FALSE;            // 消费复位请求（Consume reset request）
                _bFaultLatch := FALSE;            // 解除锁存（Release latch）
                _uErrorIdInt := 0;                // 故障码清零（Error code cleared）
                _bHoldLatch  := FALSE;            // 复位同时解除冻结（Freeze released on reset）
                _eState      := E_DL_ValveState.eIdle; // 回空闲态（Back to idle）
            END_IF
        ELSE // 锁存标志与状态不一致兜底：强制同步进故障态（Latch/state mismatch fallback）
            _eState := E_DL_ValveState.eFault;
    END_CASE
ELSE
    CASE _eState OF

        E_DL_ValveState.eIdle: // 空闲稳态：使能撤除或输出冻结
            IF bEnable AND (NOT _bHoldLatch) THEN
                _eState := E_DL_ValveState.eModulating; // 受理调节（Accept modulating）
            END_IF

        E_DL_ValveState.eModulating: // 调节中：指令整形后正常输出
            IF (NOT bEnable) OR _bHoldLatch THEN
                _eState := E_DL_ValveState.eIdle; // 使能撤除或冻结请求：输出冻结（Enable dropped or freeze requested: output frozen）
            END_IF

        ELSE // 非法状态兜底：任何越界枚举值强制锁存故障（Illegal state fallback）
            _bFaultLatch := TRUE;                 // 故障锁存（Fault latched）
            _uErrorIdInt := 16#0003_0261;         // 0003_0261 非法状态【故障级】/ Illegal state, fault level
            _eState      := E_DL_ValveState.eFault;
    END_CASE
END_IF

// ============================================================================
// 段 6｜限幅域映射与输出推导（R20：输出量纲=限幅域；冻结/故障态保持）
//      Span mapping and output derivation (output in span domain, hold in
//      frozen/fault states)
// ============================================================================
IF (_eState = E_DL_ValveState.eModulating) THEN
    _bSpanDegenerate := (ABS(_fOutMaxEff - _fOutMinEff) < 1E-9); // 跨度近零判退化（Degenerate on near-zero span）
    IF _bSpanDegenerate THEN
        _fPosOutHold := _fOutMinEff;  // 退化回退域下端（Degenerate fallback to span low）
    ELSE
        _fPosOutHold := _fOutMinEff + (_fPosCmdEff * ((_fOutMaxEff - _fOutMinEff) / 100.0)); // [%]→域线性映射（Linear mapping over span, divisor proven non-zero）
    END_IF
END_IF // 空闲/故障态不更新保持载体，输出自动冻结（Idle/fault skip update, output frozen）
fPosOutput := _fPosOutHold;           // 输出保持载体透出（Expose hold carrier）

// ============================================================================
// 段 7｜偏差报警派生与事件码优先级链（信息级瞬时每拍重算，0.15）
//      Deviation alarm derivation and event-code priority chain
// ============================================================================
_bDeviationAct := _fbTonDev.Q;        // 延时确认后激活（Active after confirmation delay）
IF (_uErrorIdInt <> 0) OR (_eState = E_DL_ValveState.eFault) THEN
    // 故障级码已锁存，信息级不覆盖（Fault-level latched, info not applied）
ELSIF _bDeviationAct THEN
    _uInfoCode := 16#0003_0112;       // 0003_0112 偏差报警激活【信息级】/ Deviation alarm active, info level
ELSIF _bSpanSwap THEN
    _uInfoCode := 16#0003_0109;       // 0003_0109 输出限幅域对调自修复【信息级】/ Span swap repair, info level
ELSIF _bClampOccur THEN
    _uInfoCode := 16#0003_0108;       // 0003_0108 设定值钳位【信息级】/ Setpoint clamped, info level
ELSE
    _uInfoCode := 0;                  // 无事件码清零（No event, code cleared）
END_IF

(*------------------------------------------------------------------------------
 * 方法: SetPosition —— 阀位指令设定 [%]，越界/非有限值拒绝返回 FALSE。
 *      Method SetPosition - position set, out-of-range or NaN returns FALSE.
 *------------------------------------------------------------------------------*)

PROPERTY eState : E_DL_ValveState
eState := _eState;            // 返回内部状态（Return internal state）

(*------------------------------------------------------------------------------
 * 属性: fPosCmd（GET）—— 当前阀位指令 [%]（钳位+死区后生效值）。
 *      Property fPosCmd (GET) - current position command [%] after shaping.
 *------------------------------------------------------------------------------*)
PROPERTY fPosCmd : REAL
fPosCmd := _fPosCmdEff;       // 返回生效指令镜像（Return effective command mirror）

(*------------------------------------------------------------------------------
 * 属性: fPosFeedback（GET）—— 阀位反馈 [%]，非有限值时保持末次有效值。
 *      Property fPosFeedback (GET) - position feedback [%], holds last valid on non-finite.
 *------------------------------------------------------------------------------*)
PROPERTY fPosFeedback : REAL
fPosFeedback := _fPosFbHold;  // 返回末次有效反馈保持值（Return last valid feedback hold value）

(*------------------------------------------------------------------------------
 * 属性: bDeviationAlarm（GET）—— 偏差报警激活中（瞬时型每拍重算）。
 *      Property bDeviationAlarm (GET) - transient deviation alarm indicator.
 *------------------------------------------------------------------------------*)
PROPERTY bDeviationAlarm : BOOL
bDeviationAlarm := _bDeviationAct; // 返回延时确认后的报警态（Return delayed-confirmed alarm state）

(*------------------------------------------------------------------------------
 * 属性: bFault（GET）—— 故障锁存指示（信息级码不置本位，0.2 公约）。
 *      Property bFault (GET) - fault latch indicator, info-level codes excluded.
 *------------------------------------------------------------------------------*)
PROPERTY bFault : BOOL
bFault := _bFaultLatch OR (_eState = E_DL_ValveState.eFault); // 显式排除信息级派生式（Explicit derived form excluding info codes）

(*------------------------------------------------------------------------------
 * 属性: uErrorId（GET）—— 末次事件码（故障级锁存优先；无故障时透出本拍
 *         信息级码，0.2/0.15 公约）。
 *      Property uErrorId (GET) - last event code (fault-level priority,
 *      transient info code shown otherwise).
 *------------------------------------------------------------------------------*)
PROPERTY uErrorId : UDINT
IF (_uErrorIdInt <> 0) OR (_eState = E_DL_ValveState.eFault) THEN
    uErrorId := _uErrorIdInt; // 故障级码优先透出（Fault-level code has priority）
ELSE
    uErrorId := _uInfoCode;   // 无故障时透出本拍信息级码（Transient info code when no fault）
END_IF
END_FUNCTION_BLOCK

(* ---- FB_DL_AnalyzerTwopointCalSeq.st ---- *)
(*==============================================================================
 * 组件 Component : FB_DL_AnalyzerTwopointCalSeq ｜ DL_Device ｜ v1.0.0 ｜ 2026-11-25
 * 功能 Function  : 水质分析仪两点标定状态机（pH/电位式电极通用）。
 *                 相序：eIdle 待机 → eZeroSettle 零液（pH 7.00）稳定判据
 *                 → eSpanSettle 标液（pH 4.00）稳定判据 → eCompute 斜率计算
 *                 → eWrite 斜率写回（域闸通过才写）→ eDone；
 *                 斜率越出接收带即走 eRollback（回滚到上一次有效斜率）并报码。
 * 边界 Boundary  : ① 稳定判据：连续 uStableCnt 拍内 |ΔmV| ≤ 0.1 mV（本文件常量），
 *                 uStableCnt=0 按 1 处理（防「零拍即稳定」的伪稳定）；
 *                 ② 同拍双窗配比约束：tZeroTmo = tSpanTmo = 120s（对称），
 *                 超时狗仅在对应相驻留时计时（R145 相驻留直驱，不叠业务补集）；
 *                 ③ 复位沿作用域三项：清锁存 / 清稳定计数与电压快照 / 迁 eIdle，
 *                 不动 _bInit；bStart 上升沿亦可重开一轮；
 *                 ④ 斜率接收带 −71.0 ~ −45.0 mV/pH（约 76%~120% 理论斜率），
 *                 越带即 eRollback：出口斜率回放上一次有效值，禁写入坏值；
 *                 ⑤ 出口 fSlopeMvPerPh 初值 = 0.0（未标定即 0，N3 安全侧），
 *                 上电不会被当作有效斜率下发。
 * 依赖 Depends   : 仅 IEC 61131-3 标准库（TON / R_TRIG / ABS）
 * 溯源 Origin    : DLF-D-WATERANA（R95 规划标签，内部原创线，无外部代码抄录）
 * 枚举归属      : E_DL_AnalyzerCalPhase 归属本文件（全库唯一属主，R264）
 * 码位分配      : 零 16# 段位范式；uErrId 常量 0 无 / 1 稳定超时 / 2 入参非有限 /
 *                 3 斜率越带（已回滚）/ 4 非法相位兜底 / 5 相位号超出映射。
 * 红线 Redline   : R1✓ R2✓ R3✓ R4✓ R5✓ R6✓（ENUM + CASE + ELSE 兜底）
 *                 R7✓（tonZero/tonSpan/rtStart/rtReset 段 0 无条件刷新） R8✓ R9✓
 *                 R14✓（无 PROPERTY） R17✓（无数组） R20✓（相位只在 CASE 内写）
 * 验收 Accept    : A1 零液 −1.0 mV 稳定 10 拍 → 标液 −178.5 mV 稳定 10 拍 →
 *                 斜率 −59.17 mV/pH，eWrite 后 bDone=TRUE；
 *                 A2 标液给 0 mV（斜率 0）→ eRollback、uErrId=3、斜率回放旧值；
 *                 A3 稳定判据长期不满足 → 120s 超时 → eFault、uErrId=1。
 *============================================================================*)

(*-----------------------------------------------------------------------------
 * 枚举: E_DL_AnalyzerCalPhase（两点标定相序）
 *----------------------------------------------------------------------------*)
TYPE E_DL_AnalyzerCalPhase :
(
    eIdle       := 0,    // 待机：等待启动沿，斜率出口保持旧值 / Idle, the slope outlet keeps the old value
    eZeroSettle := 10,   // 零液稳定判据（pH 7.00）/ Zero liquid settling with the stability criterion
    eSpanSettle := 20,   // 标液稳定判据（pH 4.00）/ Span liquid settling with the stability criterion
    eCompute    := 30,   // 斜率计算与接收带判定 / Slope computation and acceptance band check
    eWrite      := 40,   // 斜率写回 / Slope written back
    eDone       := 50,   // 完成：等待复位或重新启动 / Finished, waiting for reset or restart
    eRollback   := 60,   // 回滚：斜率越带，恢复上一次有效值 / Rollback to the last valid slope
    eFault      := 90    // 故障：超时或非有限锁存 / Fault latched by timeout or non-finite input
);
END_TYPE

FUNCTION_BLOCK FB_DL_AnalyzerTwopointCalSeq
VAR_INPUT
    bStart      : BOOL;   // 启动，上升沿开始一轮标定 [-] / Start on the rising edge
    bReset      : BOOL;   // 复位，上升沿清锁存与快照 [-] / Reset on the rising edge
    fMeasMv     : REAL;   // 电极当前电位 [mV] / Current electrode potential in millivolts
    fTempC      : REAL;   // 当前溶液温度 [°C] / Current solution temperature
    uStableCnt  : UINT;   // 稳定判据所需连续拍数，有效域 ≥ 1 [拍] / Consecutive scans required for stability
END_VAR
VAR_OUTPUT
    bDone       : BOOL;   // 本轮标定成功完成 [-] / Calibration finished successfully
    bError      : BOOL;   // 故障或回滚 [-] / Fault or rollback
    fSlopeMvPerPh : REAL; // 当前生效斜率 [mV/pH] / Slope in effect in millivolts per pH
    uErrId      : UDINT;  // 事件码锁存，0 = 无事件 [-] / Latched event code
    uPhase      : UINT;   // 相位号镜像 0/10/20/30/40/50/60/90 [-] / Phase number mirror
END_VAR
VAR
    rtStart  : R_TRIG;                                        // 启动沿实例，段 0 无条件刷新 / Start edge instance
    rtReset  : R_TRIG;                                        // 复位沿实例，段 0 无条件刷新 / Reset edge instance
    tonZero  : TON;                                           // 零液相超时狗，段 0 无条件刷新 / Zero phase watchdog
    tonSpan  : TON;                                           // 标液相超时狗，段 0 无条件刷新 / Span phase watchdog
    _eState  : E_DL_AnalyzerCalPhase := E_DL_AnalyzerCalPhase.eIdle;  // 内部相位 / Internal phase
    _bInit   : BOOL := FALSE;                                 // 首扫初始化已执行 [-] / First scan initialization done
    _bFault  : BOOL := FALSE;                                 // 故障锁存位 [-] / Latched fault bit
    _bRoll   : BOOL := FALSE;                                 // 回滚锁存位 [-] / Latched rollback bit
    _uFault  : UDINT := 0;                                    // 事件码锁存 [-] / Latched event code
    _fMvPrev : REAL := 0.0;                                   // 上一拍电位快照 [mV] / Previous potential snapshot
    _nStable : UINT := 0;                                     // 当前相内连续稳定拍数 [拍] / Consecutive stable scans in the phase
    _fMvZero : REAL := 0.0;                                   // 零液电位记录 [mV] / Recorded zero liquid potential
    _fMvSpan : REAL := 0.0;                                   // 标液电位记录 [mV] / Recorded span liquid potential
    _fSlopeNew : REAL := 0.0;                                 // 本轮新算斜率 [mV/pH] / Newly computed slope
    _fSlopeUse : REAL := 0.0;                                 // 当前生效斜率（保持量）[mV/pH] / Slope in effect
    _fSlopePrev : REAL := 0.0;                                // 上一次有效斜率（回滚目标）[mV/pH] / Last valid slope
    _bNonFin : BOOL;                                          // 入参非有限当拍量 [-] / Non-finite argument flag
    _bStableNow : BOOL;                                       // 本拍判为稳定 [-] / Stable this scan flag
    _uPhaseNew : UINT;                                        // 相位号暂存 [-] / Staged phase number
END_VAR
VAR CONSTANT
    DL_CAL_PHZERO   : REAL := 7.00;      // 零液 pH（7.00）[pH] / pH of the zero liquid
    DL_CAL_PHSPAN   : REAL := 4.00;      // 标液 pH（4.00）[pH] / pH of the span liquid
    DL_CAL_STABLEMV : REAL := 0.10;      // 稳定判据电位带 [mV] / Stability tolerance on the potential
    DL_CAL_SLO      : REAL := -71.0;     // 斜率接收带下限 [mV/pH] / Lower bound of the slope acceptance band
    DL_CAL_SHI      : REAL := -45.0;     // 斜率接收带上限 [mV/pH] / Upper bound of the slope acceptance band
    DL_CAL_TMO      : TIME := T#120S;    // 相超时时间 [ms] / Phase timeout
    DL_CAL_C_NONE   : UDINT := 0;        // 码 0：无事件 / Code zero, no event
    DL_CAL_C_TMO    : UDINT := 1;        // 码 1：稳定超时 / Code one, settling timeout
    DL_CAL_C_FIN    : UDINT := 2;        // 码 2：入参非有限 / Code two, non-finite argument
    DL_CAL_C_BAND   : UDINT := 3;        // 码 3：斜率越带已回滚 / Code three, slope out of band, rolled back
    DL_CAL_C_ILL    : UDINT := 4;        // 码 4：非法相位兜底 / Code four, illegal phase fallback
END_VAR

(* —— 段 0｜沿实例与定时器无条件每拍刷新（R7；IN 串 NOT 锁存，R145 相驻留直驱） —— *)
rtStart (CLK := bStart);
rtReset (CLK := bReset);
tonZero (IN := (_eState = E_DL_AnalyzerCalPhase.eZeroSettle) AND (NOT _bFault), PT := DL_CAL_TMO);
tonSpan (IN := (_eState = E_DL_AnalyzerCalPhase.eSpanSettle) AND (NOT _bFault), PT := DL_CAL_TMO);

(* —— 段 1｜单拍量预清零（锁存量 _bFault/_bRoll/_uFault/_nStable 不入清单，R107） —— *)
_bNonFin    := FALSE;
_bStableNow := FALSE;
_uPhaseNew  := 0;

(* —— 段 2｜首扫初始化（斜率出口落 0，N3） —— *)
IF NOT _bInit THEN
    _bInit     := TRUE;
    _bFault    := FALSE;
    _bRoll     := FALSE;
    _uFault    := DL_CAL_C_NONE;
    _fSlopeUse := 0.0;                       // 未标定：斜率 0（安全侧）
    _fSlopePrev := 0.0;
    _nStable   := 0;
    _eState    := E_DL_AnalyzerCalPhase.eIdle;
END_IF

(* —— 段 3｜复位沿处理（作用域：清锁存 / 清稳定计数与快照 / 迁相位，R311） —— *)
IF rtReset.Q THEN
    _bFault  := FALSE;                       // 作用域①：清锁存 / Scope one, clear the latches
    _bRoll   := FALSE;
    _uFault  := DL_CAL_C_NONE;
    _nStable := 0;                           // 作用域②：清计数与快照 / Scope two, clear counters
    _fMvPrev := 0.0;
    _eState  := E_DL_AnalyzerCalPhase.eIdle; // 作用域③：迁待机 / Scope three, back to idle
END_IF

(* —— 段 4｜非有限闸（覆盖参与判据的两个浮点引脚，R272） —— *)
IF (fMeasMv <> fMeasMv) OR (fTempC <> fTempC)
   OR ((fMeasMv - fMeasMv) <> (fMeasMv - fMeasMv)) THEN
    _bNonFin := TRUE;
END_IF
IF _bNonFin AND (_eState <> E_DL_AnalyzerCalPhase.eIdle) AND (NOT _bFault) THEN
    _bFault := TRUE;                         // 故障级配对（R45）
    _uFault := DL_CAL_C_FIN;
    _eState := E_DL_AnalyzerCalPhase.eFault;
END_IF

(* —— 段 5｜稳定判据（相邻拍电位差在带内即计一拍；出带即清零重计） —— *)
IF ABS(fMeasMv - _fMvPrev) <= DL_CAL_STABLEMV THEN
    _bStableNow := TRUE;
ELSE
    _nStable := 0;                           // 出带：计数清零（跨拍状态随撤销语义清零，N2）
END_IF
_fMvPrev := fMeasMv;                         // 快照唯一写入点 / Single snapshot write point

(* —— 段 6｜主状态机：八相全覆盖 + ELSE 非法相位兜底 —— *)
CASE _eState OF

E_DL_AnalyzerCalPhase.eIdle:
    IF rtStart.Q THEN
        _nStable := 0;                       // 拍 N+1 转出：进入零液稳定相
        _eState  := E_DL_AnalyzerCalPhase.eZeroSettle;
    END_IF

E_DL_AnalyzerCalPhase.eZeroSettle:
    IF _bStableNow THEN
        _nStable := _nStable + 1;
    END_IF
    IF (_nStable >= MAX(uStableCnt, 1)) THEN
        _fMvZero := fMeasMv;                 // 记录零液稳定电位
        _nStable := 0;
        _eState  := E_DL_AnalyzerCalPhase.eSpanSettle;   // 拍 N+1 转出：换标液
    ELSIF tonZero.Q THEN
        _bFault := TRUE;                     // 稳定超时：锁存（R45 配对）
        _uFault := DL_CAL_C_TMO;
        _eState := E_DL_AnalyzerCalPhase.eFault;
    END_IF

E_DL_AnalyzerCalPhase.eSpanSettle:
    IF _bStableNow THEN
        _nStable := _nStable + 1;
    END_IF
    IF (_nStable >= MAX(uStableCnt, 1)) THEN
        _fMvSpan := fMeasMv;                 // 记录标液稳定电位
        _nStable := 0;
        _eState  := E_DL_AnalyzerCalPhase.eCompute;      // 拍 N+1 转出：进入计算相
    ELSIF tonSpan.Q THEN
        _bFault := TRUE;
        _uFault := DL_CAL_C_TMO;
        _eState := E_DL_AnalyzerCalPhase.eFault;
    END_IF

E_DL_AnalyzerCalPhase.eCompute:
    (* 斜率 = ΔmV / ΔpH，ΔpH = 7.00 − 4.00 = 3.00，除子为常量非零 *)
    _fSlopeNew := (_fMvSpan - _fMvZero) / (DL_CAL_PHZERO - DL_CAL_PHSPAN);
    IF (_fSlopeNew <> _fSlopeNew) OR ((_fSlopeNew - _fSlopeNew) <> (_fSlopeNew - _fSlopeNew)) THEN
        _bFault := TRUE;                     // 计算结果非有限：故障级
        _uFault := DL_CAL_C_FIN;
        _eState := E_DL_AnalyzerCalPhase.eFault;
    ELSIF (_fSlopeNew < DL_CAL_SLO) OR (_fSlopeNew > DL_CAL_SHI) THEN
        _bRoll  := TRUE;                     // 越带：走回滚相，禁写坏值
        _uFault := DL_CAL_C_BAND;
        _eState := E_DL_AnalyzerCalPhase.eRollback;
    ELSE
        _eState := E_DL_AnalyzerCalPhase.eWrite;         // 拍 N+1 转出：写回
    END_IF

E_DL_AnalyzerCalPhase.eWrite:
    _fSlopePrev := _fSlopeUse;               // 旧值降级为回滚目标（唯一写入点）
    _fSlopeUse  := _fSlopeNew;               // 写回新斜率
    _uFault     := DL_CAL_C_NONE;
    _eState     := E_DL_AnalyzerCalPhase.eDone;

E_DL_AnalyzerCalPhase.eDone:
    IF rtStart.Q THEN
        _bRoll   := FALSE;
        _nStable := 0;
        _eState  := E_DL_AnalyzerCalPhase.eZeroSettle;   // 再次启动：重开一轮
    ELSIF rtReset.Q THEN
        _eState  := E_DL_AnalyzerCalPhase.eIdle;
    END_IF

E_DL_AnalyzerCalPhase.eRollback:
    _fSlopeUse := _fSlopePrev;               // 回滚到上一次有效斜率
    _bRoll     := TRUE;
    IF rtReset.Q OR rtStart.Q THEN
        _bRoll  := FALSE;
        _uFault := DL_CAL_C_NONE;
        _eState := E_DL_AnalyzerCalPhase.eIdle;
    END_IF

E_DL_AnalyzerCalPhase.eFault:
    _bFault := TRUE;                         // 故障相驻留：码位锁存回放（解除=bReset/bStart 沿）
    IF rtReset.Q THEN
        _uFault := DL_CAL_C_NONE;
        _eState := E_DL_AnalyzerCalPhase.eIdle;
    END_IF

ELSE
    _bFault := TRUE;                         // 非法相位兜底（R6）
    _uFault := DL_CAL_C_ILL;
    _eState := E_DL_AnalyzerCalPhase.eFault;
END_CASE

(* —— 段 7｜故障迁相闸（置于解除段之后，R274） —— *)
IF _bFault AND (_eState <> E_DL_AnalyzerCalPhase.eFault) THEN
    _eState := E_DL_AnalyzerCalPhase.eFault;
END_IF

(* —— 段 8｜统一出口段：判据位与实值单点裁决（N4 / R191） —— *)
bDone  := (_eState = E_DL_AnalyzerCalPhase.eDone);
bError := _bFault OR _bRoll;
uErrId := _uFault;
IF (_fSlopeUse <> _fSlopeUse) OR ((_fSlopeUse - _fSlopeUse) <> (_fSlopeUse - _fSlopeUse)) THEN
    fSlopeMvPerPh := 0.0;                    // 非有限兜底：斜率出口落 0（N1）
ELSE
    fSlopeMvPerPh := _fSlopeUse;
END_IF

(* 相位号镜像：单一 CASE 映射，禁多分支重复写同一状态（R20） *)
CASE _eState OF
    E_DL_AnalyzerCalPhase.eIdle:       _uPhaseNew := 0;
    E_DL_AnalyzerCalPhase.eZeroSettle: _uPhaseNew := 10;
    E_DL_AnalyzerCalPhase.eSpanSettle: _uPhaseNew := 20;
    E_DL_AnalyzerCalPhase.eCompute:    _uPhaseNew := 30;
    E_DL_AnalyzerCalPhase.eWrite:      _uPhaseNew := 40;
    E_DL_AnalyzerCalPhase.eDone:       _uPhaseNew := 50;
    E_DL_AnalyzerCalPhase.eRollback:   _uPhaseNew := 60;
    E_DL_AnalyzerCalPhase.eFault:      _uPhaseNew := 90;
ELSE
    _uPhaseNew := 90;                        // 非法相位镜像为故障号
END_CASE
uPhase := _uPhaseNew;
END_FUNCTION_BLOCK

(* ---- FB_DL_AnodizeLineTransferSeq.st ---- *)
(*==============================================================================
  Component : FB_DL_AnodizeLineTransferSeq
  Category  : DL_Device
  Type      : FB
  Complexity: C4
  VERSION   : v1.0.0
  功能      : 阳极氧化线行车转序顺控：三轴位置联动（大车 / 小车 / 升降）+ 槽位占用表互锁
  开源溯源  : 道莅原创 clean-room 自研（无外部代码引用）｜License: MIT
  边界条件  : ① 顺序闸（硬约束）：升到位（上限位）→ 才允许行走；行走到位（大车 + 小车）→ 才允许下降；
                 下降中任一轴位移信号丢失 → 同拍 E3 断能。
              ② 槽位占用表 abTankBusy 由本件唯一写入：取件相清位、放件相置位，写点各一处；
                 越界 / 占用冲突 / 非法跳槽（跨槽数 > nMaxSkipSteps 或路径中间槽被占）一律 E3。
              ③ 防双载：取件相要求吊具空载且目标槽有料；放件相要求吊具载件且目标槽空闲，
                 不满足即 E3（防丢件 / 防撞件）。方向由 _bHookLoaded 决定，无外部模式引脚。
              ④ 传感器极性义务：bPathBlockedDi / bHoistOverload 为「有障碍 / 过载」正逻辑，
                 断线失效方向（掉电无信号 = 无障碍）由 IO 适配层定义并须现场验证。
              ⑤ 默认引脚组合自证（R114）：位置与夹具类（bBridgeInPos / bTrolleyInPos / bHoistAtUpper /
                 bHoistAtLower / bClampClosed / bClampOpen）默认 FALSE，默认组合无法越过顺序闸直达放行相；
                 使能类（bEStopHealthy）默认 TRUE 与 bEnable 同族，断线由硬件安全回路保证。
              ⑥ 复位作用域（R311）：bReset 沿清 E2/E3 锁存 + 节拍 + 重试；bStop 只清 E2 与相位。
  状态机    : eIdle 待机 / eCheck 目标校验 / eLiftUp 提升到行走高度 / eTravel 大小车行走 /
              eLiftDown 下降到槽内 / eClaim 取件 / eRelease 放件 / eLiftClear 提升离槽 /
              eFault 故障停(E2) / eSafeStop 安全断能(E3)（完成结算在 eLiftClear 相内）
  自检      : R1 零 GVL ｜ R2 零物理地址 ｜ R3 纯 IEC 61131-3 ｜ R4 数组先判界 + 非有限自反判 ｜
              R6 CASE 含 ELSE ｜ R7 六 TON 两沿段 0 无条件刷新 ｜ R13 无倒序循环（单升序镜像环） ｜
              R15 定长 ARRAY，无变长数组透传 ｜ R14 无属性件
==============================================================================*)
TYPE E_DL_AtlPhase :
(
    eIdle     := 0,     (* 待机：等启动沿 / Idle, waiting for start edge *)
    eCheck    := 10,    (* 目标槽校验：越界/占用/跳槽/双载 / Target validation *)
    eLiftUp   := 20,    (* 提升到行走高度（先升后走）/ Lift to travel height *)
    eLiftDown := 40,    (* 下降到槽内（先到位再降）/ Lower into tank *)
    eTravel   := 30,    (* 大小车行走到位 / Bridge and trolley travel *)
    eClaim    := 50,    (* 取件：夹紧到位 / Claim the load *)
    eRelease  := 55,    (* 放件：松开到位 / Release the load *)
    eLiftClear:= 60,    (* 提升离槽（防撞）/ Lift clear of tank *)
    eFault    := 90,    (* 故障停待复位（E2）/ Fault stop awaiting reset, E2 *)
    eSafeStop := 95     (* 安全侧断能（E3）/ Safety energy cut, E3 *)
);
END_TYPE
TYPE E_DL_AtlCause :
(
    eNone        := 0,  (* 无异常 / No anomaly *)
    eTargetRange := 1,  (* 目标槽越界（E3）/ Target out of range, E3 *)
    eTargetSame  := 2,  (* 目标槽与当前槽相同（E3）/ Target equals current, E3 *)
    eSkipIllegal := 3,  (* 非法跳槽：跨槽数超限（E3）/ Illegal skip, E3 *)
    ePathBlocked := 4,  (* 防撞：行走路径中间槽被占（E3）/ Path blocked by occupied tank, E3 *)
    eSlotConflict:= 5,  (* 占用冲突：放件遇占用 / 取件遇空槽（E3）/ Occupancy conflict, E3 *)
    eDoubleLoad  := 6,  (* 防双载：吊具状态与任务不符（E3）/ Double-load violation, E3 *)
    eEStopOpen   := 7,  (* 急停回路断开（E3）/ E-stop circuit open, E3 *)
    eObstruct    := 8,  (* 通道障碍 / 升降过载（E3）/ Obstruction or hoist overload, E3 *)
    eLiftTmo     := 9,  (* 提升超时（E2）/ Lift-up timeout, E2 *)
    eTravelTmo   := 10, (* 行走超时（E1 记录后重试）/ Travel timeout, retried *)
    eLowerTmo    := 11, (* 下降超时（E2）/ Lower timeout, E2 *)
    eClampTmo    := 12, (* 夹取超时（E2）/ Claim timeout, E2 *)
    eOpenTmo     := 13, (* 放件超时（E2）/ Release timeout, E2 *)
    eClearTmo    := 14, (* 离槽超时（E2）/ Lift-clear timeout, E2 *)
    eRetryOver   := 15, (* 重试预算耗尽（E1 升 E2）/ Retry budget exhausted, E2 *)
    ePosBad      := 16, (* 升降位置非有限（E2）/ Hoist position non-finite, E2 *)
    eCfgBad      := 17, (* 组态非法（E2）/ Illegal configuration, E2 *)
    ePhaseBad    := 18  (* 非法相位兜底（E2）/ Illegal phase fallback, E2 *)
);
END_TYPE
TYPE E_DL_AtlGrade :
(
    eG0 := 0,           (* 无异常 / No anomaly *)
    eG1 := 1,           (* E1 可恢复重试：记录后重试，不置 bError / E1 retried, recorded only *)
    eG2 := 2,           (* E2 停机待复位 / E2 stop, awaiting reset *)
    eG3 := 3            (* E3 安全侧立即断能 / E3 immediate safety energy cut *)
);
END_TYPE

FUNCTION_BLOCK FB_DL_AnodizeLineTransferSeq
VAR_INPUT
    bStart          : BOOL := FALSE;    (* 启动沿（eIdle 入 eCheck） [-] / Start rising edge *)
    bStop           : BOOL := FALSE;    (* 中止：回 eIdle 并清 E2 锁存 [-] / Abort, clears E2 only *)
    bReset          : BOOL := FALSE;    (* 复位沿：清全部锁存 + 重试（R311） [-] / Reset edge *)
    nTargetTank     : INT := -1;        (* 目标槽号，域 0..15（-1 = 未指定） [号] / Target tank index *)
    bBridgeInPos    : BOOL := FALSE;    (* 大车到位（默认 FALSE 禁跳步） [-] / Bridge in position *)
    bTrolleyInPos   : BOOL := FALSE;    (* 小车到位（默认 FALSE 禁跳步） [-] / Trolley in position *)
    bHoistAtUpper   : BOOL := FALSE;    (* 升降上限位（行走高度） [-] / Hoist upper limit *)
    bHoistAtLower   : BOOL := FALSE;    (* 升降下限位（槽内位置） [-] / Hoist lower limit *)
    bClampClosed    : BOOL := FALSE;    (* 夹具夹紧到位 [-] / Clamp closed *)
    bClampOpen      : BOOL := FALSE;    (* 夹具松开到位 [-] / Clamp open *)
    bPathBlockedDi  : BOOL := FALSE;    (* 通道障碍（TRUE = 有障碍，正逻辑） [-] / Path obstruction *)
    bHoistOverload  : BOOL := FALSE;    (* 升降过载（TRUE = 过载，正逻辑） [-] / Hoist overload *)
    bEStopHealthy   : BOOL := TRUE;     (* 急停回路正常（使能类引脚，默认 TRUE） [-] / E-stop healthy *)
    fHoistPosMm     : LREAL := 0.0;     (* 升降实际位置（0 = 下限，向上为正） [mm] / Hoist position [mm] *)
    fHoistSafeMm    : LREAL := 500.0;   (* 行走安全高度，域 0 < v <= fHoistStrokeMm [mm] / Travel-safe height [mm] *)
    fHoistStrokeMm  : LREAL := 2000.0;  (* 升降行程上限，域 > 0 [mm] / Hoist stroke [mm] *)
    nMaxSkipSteps   : INT := 2;         (* 允许跨槽数上限，域 1..15（0 入组态闸） [槽] / Max skip [tanks] *)
    nRetryMax       : UINT := 2;        (* 行走相 E1 重试预算，域 1..9（0 入组态闸） [次] / Retry budget *)
    atPhaseTmo      : ARRAY[0..5] OF TIME := [T#60S, T#60S, T#60S, T#30S, T#30S, T#60S];   (* 超时窗 [ms]，下标 0..5 = 提升/行走/下降/夹取/放件/离槽 / Phase windows [ms] *)
    fCycleSec       : LREAL := 0.0;     (* 扫描周期（<=0 用缺省 0.01s） [s] / Scan cycle [s] *)
END_VAR
VAR_IN_OUT
    abTankBusy      : ARRAY[0..15] OF BOOL;   (* 槽位占用表（跨行车共享，写权限归本件） [-] / Tank occupancy table, written here *)
END_VAR
VAR_OUTPUT
    eState          : E_DL_AtlPhase;    (* 当前相（HMI 诊断） [-] / Present phase *)
    eCause          : E_DL_AtlCause;    (* 成因（锁存回放，R189） [-] / Latched cause playback *)
    eGrade          : E_DL_AtlGrade;    (* 异常分级出口 [-] / Exception grade outlet *)
    bError          : BOOL;             (* 故障标志（E2/E3 为 TRUE，E1 不置） [-] / Error flag *)
    bSafeCut        : BOOL;             (* 安全侧断能指令（E3 常 TRUE 至复位） [-] / Safety energy cut *)
    bHookLoaded     : BOOL;             (* 吊具载件状态（TRUE = 载件） [-] / Hook loaded state *)
    nCurrTank       : INT;              (* 行车当前槽号（-1 = 未知） [号] / Current tank index *)
    nTransferCount  : UDINT;            (* 累计转序次数（饱和） [次] / Transfer count, saturating *)
    bDone           : BOOL;             (* 单拍完成脉冲 [-] / One-scan done pulse *)
    bLiftActive     : BOOL;             (* 升降动作指示（供 IO 层驱动） [-] / Hoist action indicator *)
    bTravelActive   : BOOL;             (* 行走动作指示（供 IO 层驱动） [-] / Travel action indicator *)
    nRetryUsed      : UINT;             (* 当前相已用重试次数 [次] / Retries used in phase *)
END_VAR
VAR
    _ePhase      : E_DL_AtlPhase := E_DL_AtlPhase.eIdle;     (* 内部相（CASE 唯一写入目标） [-] / Internal phase *)
    _ePhasePrev  : E_DL_AtlPhase := E_DL_AtlPhase.eIdle;     (* 上拍相快照（相迁移后置用） [-] / Previous phase *)
    _eCause      : E_DL_AtlCause := E_DL_AtlCause.eNone;     (* 成因锁存量 [-] / Latched cause *)
    _eGrade      : E_DL_AtlGrade := E_DL_AtlGrade.eG0;       (* 分级锁存量 [-] / Latched grade *)
    _bFault      : BOOL := FALSE;       (* E2 锁存位（解除 = bReset 沿或 bStop） [-] / E2 latch *)
    _bSafeLatch  : BOOL := FALSE;       (* E3 锁存位（解除 = bReset 沿且安全恢复） [-] / E3 latch *)
    _bFaultReq   : BOOL := FALSE;       (* 单拍 E2 请求（段 1 预清，段 6 落地） [-] / One-scan E2 request *)
    _bSafeReq    : BOOL := FALSE;       (* 单拍 E3 请求（段 1 预清，段 6 落地） [-] / One-scan E3 request *)
    _bDonePulse  : BOOL := FALSE;       (* 单拍完成标志（段 1 预清） [-] / One-scan done flag *)
    _bHookLoaded : BOOL := FALSE;       (* 吊具载件内部量（分支内唯一切换） [-] / Internal hook state *)
    _bPosBad     : BOOL := FALSE;       (* 升降位置非有限当拍量 [-] / Hoist position non-finite *)
    _bCfgBad     : BOOL := FALSE;       (* 组态非法当拍量 [-] / Configuration bad *)
    _nCurr       : INT := -1;           (* 行车当前槽内部量（-1 = 未知） [号] / Internal current tank *)
    _nTarget     : INT := -1;           (* 目标槽锁存（校验通过时锁存，任务期间改目标无效） [号] / Latched target *)
    _nIdxChk     : INT := 0;            (* 相窗遍历索引（循环变量） [-] / Loop index *)
    _nRetry      : UINT := 0;           (* 当前相重试计数（相迁移后置清） [次] / Retry counter *)
    _nTransfer   : UDINT := 0;          (* 转序累计锁存（饱和） [次] / Transfer count latch *)
    _fCy         : LREAL := 0.0;        (* 当拍有效周期 [s] / Effective cycle *)
    tonLiftUp    : TON;                 (* 提升超时 / Lift-up timeout *)
    tonTravel    : TON;                 (* 行走超时（自复位，E1 可重试） / Travel timeout, self-reset *)
    tonLiftDown  : TON;                 (* 下降超时 / Lower timeout *)
    tonClaim     : TON;                 (* 取件超时 / Claim timeout *)
    tonRelease   : TON;                 (* 放件超时 / Release timeout *)
    tonLiftClear : TON;                 (* 离槽超时 / Lift-clear timeout *)
    rtStart      : R_TRIG;              (* 启动沿（段 0 无条件调用） / Start edge *)
    rtReset      : R_TRIG;              (* 复位沿（段 0 无条件调用） / Reset edge *)
END_VAR
VAR CONSTANT
    DL_ATL_TANKMAX  : INT := 15;            (* 槽号上限（ARRAY[0..15] 上界） [号] / Tank index ceiling *)
    DL_ATL_TANKCNT  : INT := 16;            (* 槽位总数（镜像取模基） [个] / Tank count *)
    DL_ATL_CYDEF    : LREAL := 0.01;        (* 缺省扫描周期 [s] / Default scan cycle [s] *)
    DL_ATL_TCNTMAX  : UDINT := 4294967295;  (* 转序计数饱和上限 [次] / Transfer count ceiling *)
    DL_ATL_RETRYTOP : UINT := 9;            (* 重试预算可配域顶 [次] / Retry configurable ceiling *)
END_VAR

(*-----------------------------------------------------------------------------
  方法 IsTankFree：槽位空闲查询（数组先判界，越界返回 FALSE 不抛错）
  契约：入参槽号越界（<0 或 >15）一律返回 FALSE，调用方须自行把它当"不可用"处理。
-----------------------------------------------------------------------------*)
METHOD PUBLIC IsTankFree : BOOL
VAR_INPUT
    nTank : INT := -1;              (* 待查槽号，域 0..15 [号] / Tank index to query *)
END_VAR

IsTankFree := FALSE;                (* 预置安全值：不可用 / Preset not-free *)
IF (nTank >= 0) AND (nTank <= DL_ATL_TANKMAX) THEN
    IF NOT abTankBusy[nTank] THEN
        IsTankFree := TRUE;         (* 界内且未占用 / In range and free *)
    END_IF
END_IF
END_METHOD

(*-----------------------------------------------------------------------------
  方法 IsPathClear：行走路径中间槽防撞校验（只扫中间槽，两端不在判据内）
  实现：先把起止槽归一为升序区间 [nLo, nHi]，再单升序循环（禁倒序循环，R13）；
        区间两端槽不属于"路径中间槽"，因此循环自 nLo+1 起、到 nHi-1 止。
-----------------------------------------------------------------------------*)
METHOD PUBLIC IsPathClear : BOOL
VAR_INPUT
    nFrom : INT := -1;              (* 起点槽号，域 0..15 [号] / Source tank *)
    nTo   : INT := -1;              (* 终点槽号，域 0..15 [号] / Destination tank *)
END_VAR
VAR
    nLo  : INT := 0;                (* 区间下界（已归一） [号] / Normalised lower bound *)
    nHi  : INT := 0;                (* 区间上界（已归一） [号] / Normalised upper bound *)
    nTmp : INT := 0;                (* 交换暂存 [号] / Swap scratch *)
    nIdx : INT := 0;                (* 升序扫描索引 [号] / Ascending index *)
END_VAR

IsPathClear := FALSE;               (* 预置不放行 / Preset not-clear *)
IF ((nFrom < 0) OR (nFrom > DL_ATL_TANKMAX)) OR ((nTo < 0) OR (nTo > DL_ATL_TANKMAX)) THEN
    IsPathClear := FALSE;           (* 端点越界：不放行 / Endpoint out of range *)
    RETURN;
END_IF
nLo := nFrom;
nHi := nTo;
IF nLo > nHi THEN
    nTmp := nLo;                    (* 归一为升序，避免倒序循环 / Normalise to ascending *)
    nLo := nHi;
    nHi := nTmp;
END_IF
IsPathClear := TRUE;                (* 默认畅通（中间槽为空集即畅通）/ Clear by default *)
FOR nIdx := nLo + 1 TO nHi - 1 DO
    IF abTankBusy[nIdx] THEN
        IsPathClear := FALSE;       (* 中间槽被占 -> 防撞拦截 / Middle tank occupied *)
    END_IF
END_FOR
END_METHOD

(*-----------------------------------------------------------------------------
  方法 NextTankIndex：从指定槽沿指定方向找下一个空闲槽（镜像取模，单升序）
  契约：nDir > 0 向后找 / nDir < 0 向前找 / nDir = 0 返回 -1（非法方向）；
        找不到空闲槽返回 -1。负模修正按 IEC 未定义行为显式补基（+16），不信平台方言。
-----------------------------------------------------------------------------*)
METHOD PUBLIC NextTankIndex : INT
VAR_INPUT
    nFrom : INT := -1;              (* 起点槽号，域 0..15 [号] / Source tank *)
    nDir  : INT := 1;               (* 方向：>0 向后 / <0 向前 [-] / Search direction *)
END_VAR
VAR
    nIdx  : INT := 0;               (* 升序步进索引 [-] / Ascending step index *)
    nCand : INT := -1;              (* 候选槽号 [号] / Candidate tank *)
END_VAR

NextTankIndex := -1;                (* 预置：未找到 / Preset not found *)
IF (nFrom < 0) OR (nFrom > DL_ATL_TANKMAX) THEN
    NextTankIndex := -1;            (* 起点越界 / Source out of range *)
    RETURN;
END_IF
IF nDir = 0 THEN
    NextTankIndex := -1;            (* 方向非法 / Illegal direction *)
    RETURN;
END_IF
FOR nIdx := 1 TO DL_ATL_TANKCNT DO
    nCand := (nFrom + nDir * nIdx) MOD DL_ATL_TANKCNT;   (* 镜像取模 / Mirror modulo *)
    IF nCand < 0 THEN
        nCand := nCand + DL_ATL_TANKCNT;                 (* 负模修正（显式补基）/ Negative modulo fix *)
    END_IF
    IF (nCand >= 0) AND (nCand <= DL_ATL_TANKMAX) THEN
        IF (NOT abTankBusy[nCand]) AND (NextTankIndex < 0) THEN
            NextTankIndex := nCand;                          (* 首个空闲槽 / First free tank *)
        END_IF
    END_IF
END_FOR
END_METHOD

(* —— 段 0：位置非有限判定 + 组态闸 + 周期派生 + 七 TON 两沿无条件刷新（R7） —— *)
_bPosBad := (fHoistPosMm <> fHoistPosMm)
         OR ((fHoistPosMm - fHoistPosMm) <> (fHoistPosMm - fHoistPosMm));   (* NaN 自反 + Inf 差值 / NaN and Inf *)
_bCfgBad := (nRetryMax = 0) OR (nRetryMax > DL_ATL_RETRYTOP)
         OR (fHoistStrokeMm <= 0.0) OR (fHoistSafeMm <= 0.0)
         OR (fHoistSafeMm > fHoistStrokeMm) OR (nMaxSkipSteps < 1) OR (nMaxSkipSteps > DL_ATL_TANKMAX);  (* 静态域闸 / Static gate *)
FOR _nIdxChk := 0 TO 5 DO
    IF atPhaseTmo[_nIdxChk] <= T#0S THEN
        _bCfgBad := TRUE;                              (* 任一相窗非正 -> 组态非法 / Non-positive window *)
    END_IF
END_FOR
IF fCycleSec > 0.0 THEN
    _fCy := fCycleSec;                                 (* 组态周期有效 / Configured cycle *)
ELSE
    _fCy := DL_ATL_CYDEF;                              (* 周期缺省兜底 / Default cycle *)
END_IF
rtStart(CLK := bStart);                                (* 启动沿，每拍必调 / Start edge every scan *)
rtReset(CLK := bReset);                                (* 复位沿，每拍必调 / Reset edge every scan *)
tonLiftUp(IN := (_ePhase = E_DL_AtlPhase.eLiftUp), PT := atPhaseTmo[0]);          (* 提升窗 / Lift window *)
tonTravel(IN := (_ePhase = E_DL_AtlPhase.eTravel) AND (NOT tonTravel.Q), PT := atPhaseTmo[1]);  (* 行走自复位窗（R188） / Travel self-reset *)
tonLiftDown(IN := (_ePhase = E_DL_AtlPhase.eLiftDown), PT := atPhaseTmo[2]);      (* 下降窗 / Lower window *)
tonClaim(IN := (_ePhase = E_DL_AtlPhase.eClaim), PT := atPhaseTmo[3]);            (* 取件窗 / Claim window *)
tonRelease(IN := (_ePhase = E_DL_AtlPhase.eRelease), PT := atPhaseTmo[4]);        (* 放件窗 / Release window *)
tonLiftClear(IN := (_ePhase = E_DL_AtlPhase.eLiftClear), PT := atPhaseTmo[5]);    (* 离槽窗 / Lift-clear window *)

(* —— 段 1：单拍量预清零（不含锁存/计数/快照量，R107）+ 相迁移后置 —— *)
_bFaultReq := FALSE;                                   (* E2 请求预清 / E2 request preset *)
_bSafeReq := FALSE;                                    (* E3 请求预清 / E3 request preset *)
_bDonePulse := FALSE;                                  (* 完成标志预清 / Done preset *)
bError := FALSE;                                       (* 故障标志预清（出口汇总） / Error preset *)
IF _ePhase <> _ePhasePrev THEN
    _nRetry := 0;                                      (* 相迁移：重试复位 / Retry reset *)
    IF _eGrade = E_DL_AtlGrade.eG1 THEN
        _eGrade := E_DL_AtlGrade.eG0;                  (* E1 记录随相推进清零 / E1 cleared on advance *)
        _eCause := E_DL_AtlCause.eNone;
    END_IF
END_IF

(* —— 段 2：E3 全局安全侧（急停 / 通道障碍 / 升降过载 / 位置非有限）——最高优先级 —— *)
IF (NOT bEStopHealthy) OR bPathBlockedDi OR bHoistOverload OR _bPosBad THEN
    IF NOT _bSafeLatch THEN
        _bSafeReq := TRUE;                             (* 请求落地位于段 6 / Landed in segment 6 *)
        IF NOT bEStopHealthy THEN
            _eCause := E_DL_AtlCause.eEStopOpen;       (* 归因：急停断开 / Cause: E-stop *)
        ELSIF _bPosBad THEN
            _eCause := E_DL_AtlCause.ePosBad;          (* 归因：位置信号非有限 / Cause: position *)
        ELSE
            _eCause := E_DL_AtlCause.eObstruct;        (* 归因：障碍或过载 / Cause: obstruction *)
        END_IF
    END_IF
END_IF

(* —— 段 3：组态闸入 E2 —— *)
IF _bCfgBad AND (NOT _bSafeLatch) AND (NOT _bFault) THEN
    _bFaultReq := TRUE;                                (* 请求落地位于段 6 / Landed in segment 6 *)
    _eCause := E_DL_AtlCause.eCfgBad;                  (* 归因：组态非法 / Cause: config *)
END_IF

(* —— 段 4：迁出链（复位沿 > 中止；作用域逐项声明 R311） —— *)
IF rtReset.Q THEN
    _bFault := FALSE;                                  (* 作用域①：清 E2 锁存 / Clear E2 *)
    IF NOT ((NOT bEStopHealthy) OR bPathBlockedDi OR bHoistOverload OR _bPosBad) THEN
        _bSafeLatch := FALSE;                          (* 作用域②：安全恢复才清 E3 / Clear E3 only if safe *)
    END_IF
    _eCause := E_DL_AtlCause.eNone;                    (* 作用域③：清成因分级 / Clear cause and grade *)
    _eGrade := E_DL_AtlGrade.eG0;
    _nRetry := 0;                                      (* 作用域④：清重试 / Clear retry *)
    IF NOT _bSafeLatch THEN
        IF (_ePhase = E_DL_AtlPhase.eFault) OR (_ePhase = E_DL_AtlPhase.eSafeStop) THEN
            _ePhase := E_DL_AtlPhase.eIdle;            (* 作用域⑤：故障相迁回待机 / Back to idle *)
        END_IF
    END_IF
ELSIF bStop AND (_ePhase <> E_DL_AtlPhase.eIdle) AND (_ePhase <> E_DL_AtlPhase.eSafeStop) THEN
    IF _ePhase = E_DL_AtlPhase.eFault THEN
        _bFault := FALSE;                              (* 中止清 E2（E3 只由复位清） / Abort clears E2 only *)
        _eCause := E_DL_AtlCause.eNone;
        _eGrade := E_DL_AtlGrade.eG0;
    END_IF
    _nRetry := 0;                                      (* 重试复位 / Retry reset *)
    _ePhase := E_DL_AtlPhase.eIdle;                    (* 回待机 / Back to idle *)
END_IF

(* —— 段 5：主状态机（顺序闸在相序与迁移判据双重固化） —— *)
CASE _ePhase OF
E_DL_AtlPhase.eIdle:
    IF rtStart.Q AND (NOT _bFault) AND (NOT _bSafeLatch) THEN
        _ePhase := E_DL_AtlPhase.eCheck;               (* 入校验相 / To check *)
    END_IF
E_DL_AtlPhase.eCheck:
    IF (nTargetTank < 0) OR (nTargetTank > DL_ATL_TANKMAX) THEN
        _eCause := E_DL_AtlCause.eTargetRange;         (* 归因：越界（E3）/ Cause: out of range *)
        _bSafeReq := TRUE;
    ELSIF (_nCurr >= 0) AND (nTargetTank = _nCurr) THEN
        _eCause := E_DL_AtlCause.eTargetSame;          (* 归因：目标等于当前（E3）/ Cause: same tank *)
        _bSafeReq := TRUE;
    ELSIF (_nCurr >= 0) AND (ABS(nTargetTank - _nCurr) > nMaxSkipSteps) THEN
        _eCause := E_DL_AtlCause.eSkipIllegal;         (* 归因：跨槽数超限（E3）/ Cause: skip too far *)
        _bSafeReq := TRUE;
    ELSIF (_nCurr >= 0) AND (NOT IsPathClear(_nCurr, nTargetTank)) THEN
        _eCause := E_DL_AtlCause.ePathBlocked;         (* 归因：路径中间槽被占（E3）/ Cause: path blocked *)
        _bSafeReq := TRUE;
    ELSIF _bHookLoaded AND (NOT IsTankFree(nTargetTank)) THEN
        _eCause := E_DL_AtlCause.eSlotConflict;        (* 放件遇占用（E3）/ Release into busy tank *)
        _bSafeReq := TRUE;
    ELSIF (NOT _bHookLoaded) AND IsTankFree(nTargetTank) THEN
        _eCause := E_DL_AtlCause.eSlotConflict;        (* 取件遇空槽（E3）/ Claim from empty tank *)
        _bSafeReq := TRUE;
    ELSIF ((NOT _bHookLoaded) AND bClampClosed) OR (_bHookLoaded AND bClampOpen) THEN
        _eCause := E_DL_AtlCause.eDoubleLoad;          (* 防双载：夹具状态与吊具记录矛盾（E3）/ Clamp state contradicts hook record *)
        _bSafeReq := TRUE;
    ELSE
        _nTarget := nTargetTank;                       (* 目标锁存：任务期间改目标无效 / Latch target *)
        _ePhase := E_DL_AtlPhase.eLiftUp;              (* 校验通过 -> 先升到位 / Valid, lift first *)
    END_IF
E_DL_AtlPhase.eLiftUp:
    IF bHoistAtUpper AND (NOT _bPosBad) THEN
        _ePhase := E_DL_AtlPhase.eTravel;              (* 升到位才允许行走 / Lift done, travel allowed *)
    ELSIF tonLiftUp.Q THEN
        _eCause := E_DL_AtlCause.eLiftTmo;             (* 归因：提升超时 / Cause: lift timeout *)
        _bFaultReq := TRUE;
    END_IF
E_DL_AtlPhase.eTravel:
    IF bBridgeInPos AND bTrolleyInPos AND (NOT bPathBlockedDi) THEN
        _ePhase := E_DL_AtlPhase.eLiftDown;            (* 两轴到位才允许下降 / Both axes in pos, lower *)
    ELSIF tonTravel.Q THEN
        IF _nRetry < nRetryMax THEN
            _nRetry := _nRetry + 1;                    (* E1：可重试，计时器自复位后重计时 / E1 retry *)
            _eGrade := E_DL_AtlGrade.eG1;
            _eCause := E_DL_AtlCause.eTravelTmo;
        ELSE
            _eCause := E_DL_AtlCause.eRetryOver;       (* 归因：重试耗尽 / Cause: retry exhausted *)
            _bFaultReq := TRUE;
        END_IF
    END_IF
E_DL_AtlPhase.eLiftDown:
    IF bHoistAtLower AND bBridgeInPos AND bTrolleyInPos THEN
        IF _bHookLoaded THEN
            _ePhase := E_DL_AtlPhase.eRelease;         (* 载件 -> 放件相 / Carrying, release *)
        ELSE
            _ePhase := E_DL_AtlPhase.eClaim;           (* 空载 -> 取件相 / Empty, claim *)
        END_IF
    ELSIF tonLiftDown.Q THEN
        _eCause := E_DL_AtlCause.eLowerTmo;            (* 归因：下降超时 / Cause: lower timeout *)
        _bFaultReq := TRUE;
    END_IF
E_DL_AtlPhase.eClaim:
    IF bClampClosed AND bHoistAtLower AND (_nTarget >= 0) AND (_nTarget <= DL_ATL_TANKMAX) THEN
        abTankBusy[_nTarget] := FALSE;              (* 占用表唯一清位点（取件）/ Single clear point *)
        _bHookLoaded := TRUE;                          (* 吊具载件 / Hook loaded *)
        _ePhase := E_DL_AtlPhase.eLiftClear;           (* 提升离槽 / Lift clear *)
    ELSIF tonClaim.Q THEN
        _eCause := E_DL_AtlCause.eClampTmo;            (* 归因：夹取超时 / Cause: claim timeout *)
        _bFaultReq := TRUE;
    END_IF
E_DL_AtlPhase.eRelease:
    IF bClampOpen AND bHoistAtLower AND (_nTarget >= 0) AND (_nTarget <= DL_ATL_TANKMAX) THEN
        abTankBusy[_nTarget] := TRUE;               (* 占用表唯一置位点（放件）/ Single set point *)
        _bHookLoaded := FALSE;                         (* 吊具空载 / Hook empty *)
        _ePhase := E_DL_AtlPhase.eLiftClear;           (* 提升离槽 / Lift clear *)
    ELSIF tonRelease.Q THEN
        _eCause := E_DL_AtlCause.eOpenTmo;             (* 归因：放件超时 / Cause: release timeout *)
        _bFaultReq := TRUE;
    END_IF
E_DL_AtlPhase.eLiftClear:
    IF bHoistAtUpper AND (NOT _bPosBad) THEN
        _nCurr := _nTarget;                            (* 当前槽更新（离槽后才确认）/ Current tank committed *)
        _bDonePulse := TRUE;                           (* 单拍完成（段 1 预清）/ One-scan done *)
        IF _nTransfer < DL_ATL_TCNTMAX THEN
            _nTransfer := _nTransfer + 1;              (* 计数推进（容量载体判上限）/ Saturating count *)
        END_IF
        _ePhase := E_DL_AtlPhase.eIdle;                (* 回待机 / Back to idle *)
    ELSIF tonLiftClear.Q THEN
        _eCause := E_DL_AtlCause.eClearTmo;            (* 归因：离槽超时 / Cause: clear timeout *)
        _bFaultReq := TRUE;
    END_IF
E_DL_AtlPhase.eFault:
    bError := TRUE;                                    (* 故障相驻留（锁存回放）/ Fault residency *)
E_DL_AtlPhase.eSafeStop:
    bError := TRUE;                                    (* 安全相驻留（锁存回放）/ Safety residency *)
ELSE
    _eCause := E_DL_AtlCause.ePhaseBad;                (* 非法相位兜底 / Illegal phase fallback *)
    _bFaultReq := TRUE;                                (* 由段 6 落地 / Landed in segment 6 *)
END_CASE

(* —— 段 6：E2/E3 请求统一落地（分支内只写成因与请求，落地仅此一处，R187/R252） —— *)
IF _bSafeReq AND (NOT _bSafeLatch) THEN
    _bSafeLatch := TRUE;                               (* E3 锁存 / Latch E3 *)
    _eGrade := E_DL_AtlGrade.eG3;                      (* 分级 E3 / Grade E3 *)
    _ePhase := E_DL_AtlPhase.eSafeStop;                (* 同步迁安全相 / Migrate *)
    bError := TRUE;                                    (* 故障标志同段置位（R45 配对）/ Error pairing *)
ELSIF _bFaultReq AND (NOT _bSafeLatch) THEN
    _bFault := TRUE;                                   (* E2 锁存 / Latch E2 *)
    _eGrade := E_DL_AtlGrade.eG2;                      (* 分级 E2 / Grade E2 *)
    _ePhase := E_DL_AtlPhase.eFault;                   (* 同步迁相（R252）/ Migrate *)
    bError := TRUE;                                    (* 故障标志同段置位（R45 配对）/ Error pairing *)
END_IF

(* —— 段 7：统一出口（电平量由 _ePhase 派生，单拍量由 _b* 标志映射） —— *)
eState := _ePhase;                                     (* 相出口 / Phase outlet *)
eCause := _eCause;                                     (* 成因回放 / Cause playback *)
eGrade := _eGrade;                                     (* 分级出口 / Grade outlet *)
bError := bError OR _bFault OR _bSafeLatch;            (* 故障标志汇总（E1 不置）/ Error summary *)
bSafeCut := _bSafeLatch;                               (* 安全断能指令 / Safety energy cut *)
bHookLoaded := _bHookLoaded;                           (* 吊具载件出口 / Hook state outlet *)
nCurrTank := _nCurr;                                   (* 当前槽出口 / Current tank outlet *)
nTransferCount := _nTransfer;                          (* 转序计数出口 / Transfer count outlet *)
bDone := _bDonePulse;                                  (* 单拍完成脉冲 / One-scan done *)
bLiftActive := (_ePhase = E_DL_AtlPhase.eLiftUp) OR (_ePhase = E_DL_AtlPhase.eLiftDown)
            OR (_ePhase = E_DL_AtlPhase.eLiftClear);   (* 升降动作指示 / Hoist indicator *)
bTravelActive := (_ePhase = E_DL_AtlPhase.eTravel);    (* 行走动作指示 / Travel indicator *)
nRetryUsed := _nRetry;                                 (* 重试占用出口 / Retry outlet *)
_ePhasePrev := _ePhase;                                (* 段末相快照 / Phase snapshot *)
END_FUNCTION_BLOCK

(* ---- FB_DL_AnodizeRinseCascadeCtrl.st ---- *)
(*
  Component : FB_DL_AnodizeRinseCascadeCtrl
  Category  : DL_Device
  Type      : FB
  Complexity: C2
  VERSION   : v1.0.0
  功能      : 逆流漂洗级联补水控制：按三级液位分级开补水阀，末级叠加电导率补水需求，末级电导超限延时报警。
  开源溯源  : 道莅原创 clean-room 自研（无外部代码引用）｜License: MIT
  边界条件  : ① 高液位须严格高于低液位、电导报警限须 > 1e-9，否则判组态非法并锁存故障；
              ② 任一液位达到高液位即强制关该级补水阀（防溢流），优先级高于电导补水；
              ③ 电导报警为延时确认型，故障锁存唯一解除路径 = bReset 上升沿。
*)
FUNCTION_BLOCK FB_DL_AnodizeRinseCascadeCtrl
VAR_INPUT
    bEnable      : BOOL;                    (* 使能电平 [-] Enable level *)
    bReset       : BOOL;                    (* 复位上升沿，清报警与故障 [-] Reset edge *)
    afLevelPct   : ARRAY[0..2] OF REAL;     (* 三级漂洗槽液位（0 为末级） [%] Rinse tank levels *)
    fCondUs      : REAL;                    (* 末级漂洗槽电导率 [μS/cm] Last stage conductivity *)
    fCondAlarmUs : REAL;                    (* 电导报警限 [μS/cm] Conductivity alarm limit *)
    fLevelLowPct : REAL;                    (* 补水启动液位 [%] Fill start level *)
    fLevelHighPct: REAL;                    (* 补水停止液位 [%] Fill stop level *)
    tCondDelay   : TIME;                    (* 电导报警确认延时 [ms] Alarm confirmation delay *)
END_VAR
VAR_OUTPUT
    abFillValve : ARRAY[0..2] OF BOOL;      (* 三级补水阀指令 [-] Fill valve commands *)
    bCondAlarm  : BOOL;                     (* 末级电导超限报警 [-] Conductivity alarm *)
    bError      : BOOL;                     (* 故障锁存标志 [-] Fault latch flag *)
    uErrId      : UDINT;                    (* 事件码，0 = 无事件 [-] Event code *)
END_VAR
VAR
    rtReset  : R_TRIG;   (* 复位沿实例，每拍无条件刷新 / Reset edge *)
    tonCond  : TON;      (* 电导报警确认计时 / Conductivity alarm timer *)
    _bFault  : BOOL;     (* 故障锁存位（锁存量） / Latched fault bit *)
    _uFault  : UDINT;    (* 故障码锁存（锁存量） / Latched fault code *)
    _bCfgBad : BOOL;     (* 组态非法当拍量 [-] Config illegal flag *)
    _bNonFin : BOOL;     (* 输入非有限当拍量 [-] Non-finite input flag *)
    nIdx     : INT;      (* 级遍历下标 [-] Stage loop index *)
    nLast    : INT;      (* 末级下标常量 [-] Last stage index *)
END_VAR
VAR CONSTANT
    DL_EPS : REAL := 1.0E-9;   (* 除零判定容差 [无量纲] Divide-by-zero tolerance *)
    DL_SEG : INT := 2;         (* 级联最高下标（三级） [-] Highest cascade index *)
END_VAR

(* —— 段 1｜每拍量预清零 + 阀门全预置（锁存量 _bFault/_uFault 不入清单） —— *)
uErrId := 16#0000_0000;
_bCfgBad := FALSE;
_bNonFin := FALSE;
nLast := DL_SEG;
FOR nIdx := 0 TO 2 DO
    IF (nIdx >= 0) AND (nIdx <= 2) THEN
        abFillValve[nIdx] := FALSE;         (* 阀门复位到关闭 [-] / Valve preset closed *)
    END_IF
END_FOR

(* —— 段 2｜非有限拦截：末级电导与三级液位逐个判（自反判 NaN，差值判 Inf） —— *)
IF (fCondUs <> fCondUs) OR ((fCondUs - fCondUs) <> 0.0)
   OR (fCondAlarmUs <> fCondAlarmUs) OR ((fCondAlarmUs - fCondAlarmUs) <> 0.0)
   OR (fLevelLowPct <> fLevelLowPct) OR ((fLevelLowPct - fLevelLowPct) <> 0.0)
   OR (fLevelHighPct <> fLevelHighPct) OR ((fLevelHighPct - fLevelHighPct) <> 0.0) THEN
    _bNonFin := TRUE;
END_IF
FOR nIdx := 0 TO 2 DO
    IF (nIdx >= 0) AND (nIdx <= 2) THEN
        IF (afLevelPct[nIdx] <> afLevelPct[nIdx])
           OR ((afLevelPct[nIdx] - afLevelPct[nIdx]) <> 0.0) THEN
            _bNonFin := TRUE;
        END_IF
    END_IF
END_FOR

(* —— 段 3｜组态闸：液位窗口上下界关系 + 电导报警限 —— *)
IF (fLevelHighPct <= fLevelLowPct) OR (fCondAlarmUs <= DL_EPS) OR (tCondDelay = T#0S) THEN
    _bCfgBad := TRUE;
END_IF
IF _bCfgBad AND (NOT _bFault) THEN
    _bFault := TRUE;
    _uFault := 16#0023_0001;                (* 故障级：组态非法 / Fault code bad config *)
END_IF
IF _bNonFin AND (NOT _bFault) THEN
    _bFault := TRUE;
    _uFault := 16#0023_0002;                (* 故障级：液位或电导非有限 / Non-finite input *)
END_IF

(* —— 段 4｜定时器每拍无条件刷新（使能挂 IN 引脚） —— *)
rtReset(CLK := bReset);
tonCond(IN := bEnable AND (NOT _bFault) AND (fCondUs > fCondAlarmUs), PT := tCondDelay);

(* —— 段 5｜复位沿：一次性清故障锁存（唯一解除路径，恒可达） —— *)
IF rtReset.Q THEN
    _bFault := FALSE;
    _uFault := 16#0000_0000;
END_IF

(* —— 段 6｜分级补水：低液位开阀；末级叠加电导超限补水；高液位强制关阀（优先级最高） —— *)
IF bEnable AND (NOT _bFault) AND (NOT _bCfgBad) AND (NOT _bNonFin) THEN
    FOR nIdx := 0 TO 2 DO
        IF (nIdx >= 0) AND (nIdx <= 2) THEN
            IF afLevelPct[nIdx] < fLevelLowPct THEN
                abFillValve[nIdx] := TRUE;  (* 低液位补水 [-] / Fill on low level *)
            END_IF
        END_IF
    END_FOR
    IF (fCondUs > fCondAlarmUs) AND (afLevelPct[nLast] < fLevelHighPct) THEN
        abFillValve[nLast] := TRUE;         (* 末级电导超限置换补水 [-] / Refresh on high conductivity *)
    END_IF
    FOR nIdx := 0 TO 2 DO
        IF (nIdx >= 0) AND (nIdx <= 2) THEN
            IF afLevelPct[nIdx] >= fLevelHighPct THEN
                abFillValve[nIdx] := FALSE; (* 高液位强制关阀，防溢流 [-] / Force close on high level *)
            END_IF
        END_IF
    END_FOR
END_IF

(* —— 段 7｜出口单点映射 —— *)
bCondAlarm := tonCond.Q AND (NOT _bFault);
bError := _bFault;
IF _bFault AND (_uFault <> 16#0000_0000) THEN
    uErrId := _uFault;                      (* 故障码锁存回放 / Latched fault replay *)
END_IF
END_FUNCTION_BLOCK
